(*
SPDX-FileCopyrightText: © 2026 Oleksandr Tiutyk <trofimich@gmail.com>
SPDX-License-Identifier: MIT
License: https://opensource.org/license/mit
*)

(*!
<summary>Describes typed generic storage and provides value access and conversion operations.</summary>
<description>
Stores a type category, address, byte size and ownership flag for externally stored data. Copying this
descriptor copies those fields, not the referenced payload. Typed access requires live storage matching the
descriptor; conversion methods do not validate its lifetime. Equals and GetHashCode share value semantics and
accept an optional borrowed IEqualityComparer. They preserve type categories, normalize floating NaN and
signed zero, and delegate nonempty OBJECT operands to the object's equality/hash pair. Neither method adds
descriptor state or takes ownership. Try methods contain exceptions and report failure without rolling back
bytes already written.
</description>
*)

{attribute 'no_explicit_call' := 'do not call this function block directly'}
FUNCTION_BLOCK GENERIC_VALUE
VAR_OUTPUT
	Address : POINTER TO BYTE;
	Size : ULINT;
	TypeClass : GENERIC_TYPE_CLASS;
	IsMemoryOwner : BOOL;
END_VAR

(*!
<summary>Returns a borrowed system descriptor for this generic value.</summary>
<description>
Does not copy the payload or transfer ownership. Size above SignedInt32.MAX_VALUE raises
ArgumentOutOfRangeException; type mapping exceptions propagate. The caller keeps the described storage alive
while using the result. Descendants cannot override this descriptor operation; customize value equality
through IEqualityComparer or the stored object equality contract.
</description>
*)
METHOD FINAL AsAnyType : __SYSTEM.AnyType
AsAnyType := SystemAnyTypes.CreateAnyTypeByGenericValue(genericValue := THIS^);
END_METHOD

(*!
<summary>Reads a Boolean or converts an integer to FALSE for zero and TRUE for any nonzero value.</summary>
<description>
Requires live storage matching the descriptor. Signed and unsigned integers are read at their full width,
including BYTE, WORD, DWORD and LWORD representations. Other categories throw
GenericConversionNotSupportedException. Stored data and ownership are unchanged. Descendants cannot override
this descriptor operation; customize value equality through IEqualityComparer or the stored object equality
contract.
</description>
*)
METHOD FINAL AsBool : BOOL
VAR
	universalPointer : UNIVERSAL_POINTER;
END_VAR
universalPointer.AsByte := Address;

CASE TypeClass OF
	GENERIC_TYPE_CLASS.BOOLEAN:
		AsBool := universalPointer.AsBool^;
		RETURN;

	GENERIC_TYPE_CLASS.INT_8, GENERIC_TYPE_CLASS.INT_16, GENERIC_TYPE_CLASS.INT_32, GENERIC_TYPE_CLASS.INT_64:
		AsBool := AsLInt() <> 0;
		RETURN;

	GENERIC_TYPE_CLASS.UINT_8, GENERIC_TYPE_CLASS.UINT_16, GENERIC_TYPE_CLASS.UINT_32, GENERIC_TYPE_CLASS.UINT_64:
		AsBool := AsULInt() <> 0;
		RETURN;
END_CASE

Exceptions.ThrowGenericConversionNotSupported(
		sourceNamespaceName := NamespaceName,
		sourceClassName := ClassName,
		sourcePOUName := __POUNAME(),
		sourcePosition := __POSITION(),
		sourceDataType := TypeClass,
		targetDataType := GENERIC_TYPE_CLASS.BOOLEAN
	);
END_METHOD

(*!
<summary>Reads or converts an integer representation when the value fits the result.</summary>
<description>
Requires live storage matching the descriptor. For supported integer types, FALSE accepts the actual value
only when it fits the result range; bounds are checked before narrowing or changing signedness. TRUE permits
the native conversion even outside that range. Unsupported types or rejected values raise
GenericConversionNotSupportedException. Existing BOOLEAN byte-view behavior is retained. Stored data and
ownership are unchanged; no dynamic allocation is needed for successful conversion. Descendants cannot
override this descriptor operation; customize value equality through IEqualityComparer or the stored object
equality contract.
</description>
*)
//!<param name="allowTypeCastWithDataLoss">
//! Allows native conversion when the actual value is outside the result range; overflow behavior follows
//! TwinCAT.
//! </param>
METHOD FINAL AsByte : BYTE
VAR_INPUT
	allowTypeCastWithDataLoss : BOOL := FALSE;
END_VAR
VAR
	universalPointer : UNIVERSAL_POINTER;
END_VAR
universalPointer.AsByte := Address;

CASE TypeClass OF
	GENERIC_TYPE_CLASS.BOOLEAN, GENERIC_TYPE_CLASS.UINT_8:
		 AsByte := universalPointer.AsByte^;
		 RETURN;

	GENERIC_TYPE_CLASS.UINT_16:
		IF allowTypeCastWithDataLoss OR_ELSE (TO_ULINT(universalPointer.AsWord^) <= TO_ULINT(UnsignedInt8.MAX_VALUE)) THEN
			AsByte := TO_BYTE(universalPointer.AsWord^);
			RETURN;
		END_IF

	GENERIC_TYPE_CLASS.UINT_32:
		IF allowTypeCastWithDataLoss OR_ELSE (TO_ULINT(universalPointer.AsDWord^) <= TO_ULINT(UnsignedInt8.MAX_VALUE)) THEN
			AsByte := TO_BYTE(universalPointer.AsDWord^);
			RETURN;
		END_IF

	GENERIC_TYPE_CLASS.UINT_64:
		IF allowTypeCastWithDataLoss OR_ELSE (TO_ULINT(universalPointer.AsLWord^) <= TO_ULINT(UnsignedInt8.MAX_VALUE)) THEN
			AsByte := TO_BYTE(universalPointer.AsLWord^);
			RETURN;
		END_IF

	GENERIC_TYPE_CLASS.INT_8:
		IF allowTypeCastWithDataLoss OR_ELSE (TO_LINT(universalPointer.AsSInt^) >= TO_LINT(UnsignedInt8.MIN_VALUE)) THEN
			AsByte := TO_BYTE(universalPointer.AsSInt^);
			RETURN;
		END_IF

	GENERIC_TYPE_CLASS.INT_16:
		IF allowTypeCastWithDataLoss
			OR_ELSE (TO_LINT(universalPointer.AsInt^) >= TO_LINT(UnsignedInt8.MIN_VALUE)
				AND_THEN TO_LINT(universalPointer.AsInt^) <= TO_LINT(UnsignedInt8.MAX_VALUE))
		THEN
			AsByte := TO_BYTE(universalPointer.AsInt^);
			RETURN;
		END_IF

	GENERIC_TYPE_CLASS.INT_32:
		IF allowTypeCastWithDataLoss
			OR_ELSE (TO_LINT(universalPointer.AsDInt^) >= TO_LINT(UnsignedInt8.MIN_VALUE)
				AND_THEN TO_LINT(universalPointer.AsDInt^) <= TO_LINT(UnsignedInt8.MAX_VALUE))
		THEN
			AsByte := TO_BYTE(universalPointer.AsDInt^);
			RETURN;
		END_IF

	GENERIC_TYPE_CLASS.INT_64:
		IF allowTypeCastWithDataLoss
			OR_ELSE (TO_LINT(universalPointer.AsLInt^) >= TO_LINT(UnsignedInt8.MIN_VALUE)
				AND_THEN TO_LINT(universalPointer.AsLInt^) <= TO_LINT(UnsignedInt8.MAX_VALUE))
		THEN
			AsByte := TO_BYTE(universalPointer.AsLInt^);
			RETURN;
		END_IF
END_CASE

Exceptions.ThrowGenericConversionNotSupported(
		sourceNamespaceName := NamespaceName,
		sourceClassName := ClassName,
		sourcePOUName := __POUNAME(),
		sourcePosition := __POSITION(),
		sourceDataType := TypeClass,
		targetDataType := GENERIC_TYPE_CLASS.UINT_8
	);
END_METHOD

(*!
<summary>Reads or converts a supported generic value to DATE.</summary>
<description>
Requires live storage matching the descriptor. INT_32, UINT_32, INT_64 and UINT_64 are counts of seconds since
the epoch; DATE_AND_TIME_32 is a calendar timestamp. Numeric inputs must fit DateAndTimes.MIN_VALUE/MAX_VALUE
even with TRUE. LDATE is checked as signed nanoseconds against the same limits widened to LDT before
narrowing. For these inputs, FALSE accepts only midnight; TRUE discards the time of day. The result of these
conversions has no hidden time remainder. Rejected or unsupported conversions raise
GenericConversionNotSupportedException. DATE_32 is read directly. A valid calendar LDATE within the DATE range
is accepted with either flag; a hidden time remainder requires TRUE and is explicitly removed. Stored data and
ownership are unchanged. Descendants cannot override this descriptor operation; customize value equality
through IEqualityComparer or the stored object equality contract.
</description>
*)
//!<param name="allowTypeCastWithDataLoss">
//! Allows discarding the time of day from numeric, DT and LDATE inputs; does not permit numeric or LDATE
//! range overflow.
//! </param>
METHOD FINAL AsDate : DATE
VAR_INPUT
	allowTypeCastWithDataLoss : BOOL := FALSE;
END_VAR
VAR
	universalPointer : UNIVERSAL_POINTER;

	secondsSinceMidnight : UDINT;
END_VAR
universalPointer.AsByte := Address;

CASE TypeClass OF
	GENERIC_TYPE_CLASS.DATE_32: 
		 AsDate := universalPointer.AsDate^;
		 RETURN;		 

	GENERIC_TYPE_CLASS.INT_32:
		IF universalPointer.AsDInt^ >= TO_LINT(DateAndTimes.MIN_VALUE) THEN
			secondsSinceMidnight := TO_UDINT(universalPointer.AsDInt^) MOD Times.SECONDS_PER_DAY;

			IF allowTypeCastWithDataLoss
				OR_ELSE secondsSinceMidnight = 0
			THEN
				AsDate := TO_DATE(TO_UDINT(universalPointer.AsDInt^) - secondsSinceMidnight);
				RETURN;
			END_IF
		END_IF

	GENERIC_TYPE_CLASS.UINT_32, GENERIC_TYPE_CLASS.DATE_AND_TIME_32:
		secondsSinceMidnight := TO_UDINT(universalPointer.AsUDInt^) MOD Times.SECONDS_PER_DAY;

		IF allowTypeCastWithDataLoss
			OR_ELSE secondsSinceMidnight = 0
		THEN
			AsDate := TO_DATE(TO_UDINT(universalPointer.AsUDInt^) - secondsSinceMidnight);
			RETURN;
		END_IF

	GENERIC_TYPE_CLASS.INT_64:
		IF universalPointer.AsLInt^ >= TO_LINT(DateAndTimes.MIN_VALUE) AND_THEN universalPointer.AsLInt^ <= TO_LINT(DateAndTimes.MAX_VALUE) THEN
			secondsSinceMidnight := TO_UDINT(universalPointer.AsLInt^) MOD Times.SECONDS_PER_DAY;

			IF allowTypeCastWithDataLoss
				OR_ELSE secondsSinceMidnight = 0
			THEN
				AsDate := TO_DATE(TO_UDINT(universalPointer.AsLInt^) - secondsSinceMidnight);
				RETURN;
			END_IF
		END_IF

	GENERIC_TYPE_CLASS.UINT_64:
		IF universalPointer.AsULInt^ <= TO_ULINT(DateAndTimes.MAX_VALUE) THEN
			secondsSinceMidnight := TO_UDINT(universalPointer.AsULInt^) MOD Times.SECONDS_PER_DAY;

			IF allowTypeCastWithDataLoss
				OR_ELSE secondsSinceMidnight = 0
			THEN
				AsDate := TO_DATE(TO_UDINT(universalPointer.AsULInt^) - secondsSinceMidnight);
				RETURN;
			END_IF
		END_IF

	GENERIC_TYPE_CLASS.DATE_64:
		IF universalPointer.AsLInt^ >= TO_LINT(TO_LDT(DateAndTimes.MIN_VALUE))
			AND_THEN universalPointer.AsLInt^ <= TO_LINT(TO_LDT(DateAndTimes.MAX_VALUE)) THEN
			IF allowTypeCastWithDataLoss OR_ELSE universalPointer.AsLInt^ MOD TO_LINT(LongTimes.ONE_DAY) = 0 THEN
				// Remove the time in nanoseconds before converting whole seconds to DATE.
				AsDate := TO_DATE((universalPointer.AsLInt^ - universalPointer.AsLInt^ MOD TO_LINT(LongTimes.ONE_DAY))
					/ TO_LINT(LongTimes.ONE_SECOND));
				RETURN;
			END_IF
		END_IF
END_CASE

Exceptions.ThrowGenericConversionNotSupported(
		sourceNamespaceName := NamespaceName,
		sourceClassName := ClassName,
		sourcePOUName := __POUNAME(),
		sourcePosition := __POSITION(),
		sourceDataType := TypeClass,
		targetDataType := GENERIC_TYPE_CLASS.DATE_32
	);
END_METHOD

(*!
<summary>Reads or converts a supported generic value to DATE_AND_TIME.</summary>
<description>
Requires live storage matching the descriptor. For DATE_AND_TIME_64, FALSE requires a timestamp within the DT
range and an exact whole number of seconds. Signed nanoseconds are checked before narrowing. TRUE uses native
TO_DT without these checks; out-of-range behavior depends on the runtime and may raise an exception. Rejected
or unsupported conversions raise GenericConversionNotSupportedException. Numeric inputs are seconds since the
epoch. With FALSE, signed inputs must be nonnegative and 64-bit inputs must fit the DT range; TRUE passes the
original signed or unsigned value to native TO_DT. DATE_32 and DATE_AND_TIME_32 retain their direct conversion
paths. Stored data and ownership are unchanged. Descendants cannot override this descriptor operation;
customize value equality through IEqualityComparer or the stored object equality contract.
</description>
*)
//!<param name="allowTypeCastWithDataLoss">
//! Allows loss of precision or range in LDT to DT conversion and native numeric conversions outside the DT
//! range.
//! </param>
METHOD FINAL AsDateAndTime : DATE_AND_TIME
VAR_INPUT
	allowTypeCastWithDataLoss : BOOL := FALSE;
END_VAR
VAR
	universalPointer : UNIVERSAL_POINTER;
END_VAR
universalPointer.AsByte := Address;

CASE TypeClass OF
	GENERIC_TYPE_CLASS.DATE_AND_TIME_32:
		 AsDateAndTime := universalPointer.AsDateAndTime^;
		 RETURN;

	GENERIC_TYPE_CLASS.UINT_32:
		 AsDateAndTime := TO_DT(universalPointer.AsUDInt^);
		 RETURN;
		
	GENERIC_TYPE_CLASS.DATE_32:
		 AsDateAndTime := TO_DT(universalPointer.AsDate^);
		 RETURN;
	GENERIC_TYPE_CLASS.DATE_AND_TIME_64:
		IF allowTypeCastWithDataLoss OR_ELSE (
			universalPointer.AsLInt^ >= TO_LINT(TO_LDT(DateAndTimes.MIN_VALUE))
			AND_THEN universalPointer.AsLInt^ <= TO_LINT(TO_LDT(DateAndTimes.MAX_VALUE))
			AND_THEN universalPointer.AsLInt^ MOD TO_LINT(LongTimes.ONE_SECOND) = 0) THEN
			AsDateAndTime := TO_DT(universalPointer.AsLDateAndTime^);
			RETURN;
		END_IF

	GENERIC_TYPE_CLASS.INT_32:
		IF allowTypeCastWithDataLoss OR_ELSE universalPointer.AsDInt^ >= TO_LINT(DateAndTimes.MIN_VALUE) THEN
			AsDateAndTime := TO_DT(universalPointer.AsDInt^);
			RETURN;
		END_IF

	GENERIC_TYPE_CLASS.INT_64:
		IF allowTypeCastWithDataLoss OR_ELSE (
			universalPointer.AsLInt^ >= TO_LINT(DateAndTimes.MIN_VALUE)
			AND_THEN universalPointer.AsLInt^ <= TO_LINT(DateAndTimes.MAX_VALUE)) THEN
			AsDateAndTime := TO_DT(universalPointer.AsLInt^);
			RETURN;
		END_IF

	GENERIC_TYPE_CLASS.UINT_64:
		IF allowTypeCastWithDataLoss OR_ELSE universalPointer.AsULInt^ <= TO_ULINT(DateAndTimes.MAX_VALUE) THEN
			AsDateAndTime := TO_DT(universalPointer.AsULInt^);
			RETURN;
		END_IF
END_CASE

Exceptions.ThrowGenericConversionNotSupported(
		sourceNamespaceName := NamespaceName,
		sourceClassName := ClassName,
		sourcePOUName := __POUNAME(),
		sourcePosition := __POSITION(),
		sourceDataType := TypeClass,
		targetDataType := GENERIC_TYPE_CLASS.DATE_AND_TIME_32
	);
END_METHOD

(*!
<summary>Reads or converts an integer representation when the value fits the result.</summary>
<description>
Requires live storage matching the descriptor. For supported integer types, FALSE accepts the actual value
only when it fits the result range; bounds are checked before narrowing or changing signedness. TRUE permits
the native conversion even outside that range. Unsupported types or rejected values raise
GenericConversionNotSupportedException. Existing BOOLEAN byte-view behavior is retained. Stored data and
ownership are unchanged; no dynamic allocation is needed for successful conversion. Descendants cannot
override this descriptor operation; customize value equality through IEqualityComparer or the stored object
equality contract.
</description>
*)
//!<param name="allowTypeCastWithDataLoss">
//! Allows native conversion when the actual value is outside the result range; overflow behavior follows
//! TwinCAT.
//! </param>
METHOD FINAL AsDInt : DINT
VAR_INPUT
	allowTypeCastWithDataLoss : BOOL := FALSE;
END_VAR
VAR
	universalPointer : UNIVERSAL_POINTER;
END_VAR
universalPointer.AsByte := Address;

CASE TypeClass OF
	GENERIC_TYPE_CLASS.BOOLEAN, GENERIC_TYPE_CLASS.UINT_8:
		 AsDInt := TO_DINT(universalPointer.AsByte^);
		 RETURN;
		
	GENERIC_TYPE_CLASS.UINT_16:
		 AsDInt := TO_DINT(universalPointer.AsWord^);
		 RETURN;

	GENERIC_TYPE_CLASS.INT_8: 
		 AsDInt := TO_DINT(universalPointer.AsSInt^);
		 RETURN;
		 
	GENERIC_TYPE_CLASS.INT_16: 
		 AsDInt := TO_DINT(universalPointer.AsInt^);
		 RETURN;
		 
	GENERIC_TYPE_CLASS.INT_32: 
		 AsDInt := universalPointer.AsDInt^;
		 RETURN;

	GENERIC_TYPE_CLASS.UINT_32:
		IF allowTypeCastWithDataLoss OR_ELSE (TO_ULINT(universalPointer.AsDWord^) <= TO_ULINT(SignedInt32.MAX_VALUE)) THEN
			AsDInt := TO_DINT(universalPointer.AsDWord^);
			RETURN;
		END_IF

	GENERIC_TYPE_CLASS.UINT_64:
		IF allowTypeCastWithDataLoss OR_ELSE (TO_ULINT(universalPointer.AsLWord^) <= TO_ULINT(SignedInt32.MAX_VALUE)) THEN
			AsDInt := TO_DINT(universalPointer.AsLWord^);
			RETURN;
		END_IF

	GENERIC_TYPE_CLASS.INT_64:
		IF allowTypeCastWithDataLoss
			OR_ELSE (TO_LINT(universalPointer.AsLInt^) >= TO_LINT(SignedInt32.MIN_VALUE)
				AND_THEN TO_LINT(universalPointer.AsLInt^) <= TO_LINT(SignedInt32.MAX_VALUE))
		THEN
			AsDInt := TO_DINT(universalPointer.AsLInt^);
			RETURN;
		END_IF
END_CASE

Exceptions.ThrowGenericConversionNotSupported(
		sourceNamespaceName := NamespaceName,
		sourceClassName := ClassName,
		sourcePOUName := __POUNAME(),
		sourcePosition := __POSITION(),
		sourceDataType := TypeClass,
		targetDataType := GENERIC_TYPE_CLASS.INT_32
	);
END_METHOD

(*!
<summary>Reads or converts an integer representation when the value fits the result.</summary>
<description>
Requires live storage matching the descriptor. For supported integer types, FALSE accepts the actual value
only when it fits the result range; bounds are checked before narrowing or changing signedness. TRUE permits
the native conversion even outside that range. Unsupported types or rejected values raise
GenericConversionNotSupportedException. Existing BOOLEAN byte-view behavior is retained. Stored data and
ownership are unchanged; no dynamic allocation is needed for successful conversion. Descendants cannot
override this descriptor operation; customize value equality through IEqualityComparer or the stored object
equality contract.
</description>
*)
//!<param name="allowTypeCastWithDataLoss">
//! Allows native conversion when the actual value is outside the result range; overflow behavior follows
//! TwinCAT.
//! </param>
METHOD FINAL AsDWord : DWORD
VAR_INPUT
	allowTypeCastWithDataLoss : BOOL := FALSE;
END_VAR
VAR
	universalPointer : UNIVERSAL_POINTER;
END_VAR
universalPointer.AsByte := Address;

CASE TypeClass OF
	GENERIC_TYPE_CLASS.BOOLEAN, GENERIC_TYPE_CLASS.UINT_8:
		 AsDWord := TO_DWORD(universalPointer.AsByte^);
		 RETURN;
		 
	GENERIC_TYPE_CLASS.UINT_16:
		 AsDWord := TO_DWORD(universalPointer.AsWord^);
		 RETURN;
 
	GENERIC_TYPE_CLASS.UINT_32: 
		 AsDWord := universalPointer.AsDWord^;
		 RETURN;

	GENERIC_TYPE_CLASS.UINT_64:
		IF allowTypeCastWithDataLoss OR_ELSE (TO_ULINT(universalPointer.AsLWord^) <= TO_ULINT(UnsignedInt32.MAX_VALUE)) THEN
			AsDWord := TO_DWORD(universalPointer.AsLWord^);
			RETURN;
		END_IF

	GENERIC_TYPE_CLASS.INT_8:
		IF allowTypeCastWithDataLoss OR_ELSE (TO_LINT(universalPointer.AsSInt^) >= TO_LINT(UnsignedInt32.MIN_VALUE)) THEN
			AsDWord := TO_DWORD(universalPointer.AsSInt^);
			RETURN;
		END_IF

	GENERIC_TYPE_CLASS.INT_16:
		IF allowTypeCastWithDataLoss OR_ELSE (TO_LINT(universalPointer.AsInt^) >= TO_LINT(UnsignedInt32.MIN_VALUE)) THEN
			AsDWord := TO_DWORD(universalPointer.AsInt^);
			RETURN;
		END_IF

	GENERIC_TYPE_CLASS.INT_32:
		IF allowTypeCastWithDataLoss OR_ELSE (TO_LINT(universalPointer.AsDInt^) >= TO_LINT(UnsignedInt32.MIN_VALUE)) THEN
			AsDWord := TO_DWORD(universalPointer.AsDInt^);
			RETURN;
		END_IF

	GENERIC_TYPE_CLASS.INT_64:
		IF allowTypeCastWithDataLoss
			OR_ELSE (TO_LINT(universalPointer.AsLInt^) >= TO_LINT(UnsignedInt32.MIN_VALUE)
				AND_THEN TO_LINT(universalPointer.AsLInt^) <= TO_LINT(UnsignedInt32.MAX_VALUE))
		THEN
			AsDWord := TO_DWORD(universalPointer.AsLInt^);
			RETURN;
		END_IF
END_CASE

Exceptions.ThrowGenericConversionNotSupported(
		sourceNamespaceName := NamespaceName,
		sourceClassName := ClassName,
		sourcePOUName := __POUNAME(),
		sourcePosition := __POSITION(),
		sourceDataType := TypeClass,
		targetDataType := GENERIC_TYPE_CLASS.UINT_32
	);
END_METHOD

(*!
<summary>Reads or converts an integer representation when the value fits the result.</summary>
<description>
Requires live storage matching the descriptor. For supported integer types, FALSE accepts the actual value
only when it fits the result range; bounds are checked before narrowing or changing signedness. TRUE permits
the native conversion even outside that range. Unsupported types or rejected values raise
GenericConversionNotSupportedException. Existing BOOLEAN byte-view behavior is retained. Stored data and
ownership are unchanged; no dynamic allocation is needed for successful conversion. Descendants cannot
override this descriptor operation; customize value equality through IEqualityComparer or the stored object
equality contract.
</description>
*)
//!<param name="allowTypeCastWithDataLoss">
//! Allows native conversion when the actual value is outside the result range; overflow behavior follows
//! TwinCAT.
//! </param>
METHOD FINAL AsInt : INT
VAR_INPUT
	allowTypeCastWithDataLoss : BOOL := FALSE;
END_VAR
VAR
	universalPointer : UNIVERSAL_POINTER;
END_VAR
universalPointer.AsByte := Address;

CASE TypeClass OF
	GENERIC_TYPE_CLASS.BOOLEAN, GENERIC_TYPE_CLASS.UINT_8:
		 AsInt := TO_INT(universalPointer.AsByte^);
		 RETURN;

	GENERIC_TYPE_CLASS.INT_8: 
		 AsInt := TO_INT(universalPointer.AsSInt^);
		 RETURN;
			 
	GENERIC_TYPE_CLASS.INT_16: 
		 AsInt := universalPointer.AsInt^;
		 RETURN;

	GENERIC_TYPE_CLASS.UINT_16:
		IF allowTypeCastWithDataLoss OR_ELSE (TO_ULINT(universalPointer.AsWord^) <= TO_ULINT(SignedInt16.MAX_VALUE)) THEN
			AsInt := TO_INT(universalPointer.AsWord^);
			RETURN;
		END_IF

	GENERIC_TYPE_CLASS.UINT_32:
		IF allowTypeCastWithDataLoss OR_ELSE (TO_ULINT(universalPointer.AsDWord^) <= TO_ULINT(SignedInt16.MAX_VALUE)) THEN
			AsInt := TO_INT(universalPointer.AsDWord^);
			RETURN;
		END_IF

	GENERIC_TYPE_CLASS.UINT_64:
		IF allowTypeCastWithDataLoss OR_ELSE (TO_ULINT(universalPointer.AsLWord^) <= TO_ULINT(SignedInt16.MAX_VALUE)) THEN
			AsInt := TO_INT(universalPointer.AsLWord^);
			RETURN;
		END_IF

	GENERIC_TYPE_CLASS.INT_32:
		IF allowTypeCastWithDataLoss
			OR_ELSE (TO_LINT(universalPointer.AsDInt^) >= TO_LINT(SignedInt16.MIN_VALUE)
				AND_THEN TO_LINT(universalPointer.AsDInt^) <= TO_LINT(SignedInt16.MAX_VALUE))
		THEN
			AsInt := TO_INT(universalPointer.AsDInt^);
			RETURN;
		END_IF

	GENERIC_TYPE_CLASS.INT_64:
		IF allowTypeCastWithDataLoss
			OR_ELSE (TO_LINT(universalPointer.AsLInt^) >= TO_LINT(SignedInt16.MIN_VALUE)
				AND_THEN TO_LINT(universalPointer.AsLInt^) <= TO_LINT(SignedInt16.MAX_VALUE))
		THEN
			AsInt := TO_INT(universalPointer.AsLInt^);
			RETURN;
		END_IF
END_CASE

Exceptions.ThrowGenericConversionNotSupported(
		sourceNamespaceName := NamespaceName,
		sourceClassName := ClassName,
		sourcePOUName := __POUNAME(),
		sourcePosition := __POSITION(),
		sourceDataType := TypeClass,
		targetDataType := GENERIC_TYPE_CLASS.INT_16
	);
END_METHOD

(*!
<summary>Returns a borrowed IObject view of object storage.</summary>
<description>
Requires OBJECT TypeClass; other tags raise GenericConversionNotSupportedException. A null address returns a
null interface; a nonnull address must identify a live compatible object. Does not clone or transfer
ownership. Descendants cannot override this descriptor operation; customize value equality through
IEqualityComparer or the stored object equality contract.
</description>
*)
METHOD FINAL AsIObject : IObject
VAR
	objectPointer : POINTER TO Object;

END_VAR
IF TypeClass = GENERIC_TYPE_CLASS.OBJECT THEN
	objectPointer := Address;
	
	IF objectPointer <> 0 THEN
		__QUERYINTERFACE(objectPointer^, AsIObject);						
	END_IF
ELSE	
	Exceptions.ThrowGenericConversionNotSupported(
		sourceNamespaceName := NamespaceName,
		sourceClassName := ClassName,
		sourcePOUName := __POUNAME(),
		sourcePosition := __POSITION(),
		sourceDataType := TypeClass,
		targetDataType := GENERIC_TYPE_CLASS.OBJECT
	);		
END_IF
END_METHOD

(*!
<summary>Reads or converts a supported generic value to LDATE.</summary>
<description>
Requires live storage matching the descriptor. DATE_AND_TIME_32 and DATE_AND_TIME_64 are treated as calendar
timestamps. INT_64 and UINT_64 are signed and unsigned counts of nanoseconds since the epoch. UINT_64 values
above LongDateAndTimes.MAX_VALUE are rejected even with TRUE. Numeric inputs follow calendar normalization:
FALSE accepts only midnight; TRUE discards the time of day. The results have no hidden time remainder. LDT
normalization uses signed nanoseconds and rounds down to midnight, including before the epoch. The first
partial LDT day (1677-09-21) is rejected even with TRUE because its midnight cannot be represented in LDATE;
the range check precedes subtraction. Rejected or unsupported conversions raise
GenericConversionNotSupportedException. DATE_64 is read directly and DATE_32 uses native widening; these paths
do not normalize hidden time components. Stored data and ownership are unchanged. Descendants cannot override
this descriptor operation; customize value equality through IEqualityComparer or the stored object equality
contract.
</description>
*)
//!<param name="allowTypeCastWithDataLoss">
//! Allows discarding the time of day from DT, LDT and numeric nanosecond counts; does not permit a midnight
//! outside the LDATE range.
//! </param>
METHOD FINAL AsLDate : LDATE
VAR_INPUT
	allowTypeCastWithDataLoss : BOOL := FALSE;
END_VAR
VAR
	universalPointer : UNIVERSAL_POINTER;

	secondsSinceMidnight : UDINT;
	nanosecondsSinceMidnight : LINT;
END_VAR
universalPointer.AsByte := Address;

CASE TypeClass OF
	GENERIC_TYPE_CLASS.DATE_64: 
		 AsLDate := universalPointer.AsLDate^;
		 RETURN;		 

	GENERIC_TYPE_CLASS.DATE_32: 
		 AsLDate := TO_LDATE(universalPointer.AsDate^);
		 RETURN;
	GENERIC_TYPE_CLASS.UINT_64:
		IF universalPointer.AsULInt^ <= TO_ULINT(LongDateAndTimes.MAX_VALUE) THEN
			nanosecondsSinceMidnight := TO_LINT(universalPointer.AsULInt^ MOD TO_ULINT(LongTimes.ONE_DAY));

			IF allowTypeCastWithDataLoss
				OR_ELSE nanosecondsSinceMidnight = 0
			THEN
				AsLDate := TO_LDATE(universalPointer.AsULInt^ - TO_ULINT(nanosecondsSinceMidnight));
				RETURN;
			END_IF
		END_IF

	GENERIC_TYPE_CLASS.DATE_AND_TIME_32:
		secondsSinceMidnight := TO_UDINT(universalPointer.AsDateAndTime^) MOD Times.SECONDS_PER_DAY;

		IF allowTypeCastWithDataLoss
			OR_ELSE secondsSinceMidnight = 0
		THEN
			AsLDate := TO_LDATE(TO_DT(TO_UDINT(universalPointer.AsDateAndTime^) - secondsSinceMidnight));
			RETURN;
		END_IF

	GENERIC_TYPE_CLASS.DATE_AND_TIME_64, GENERIC_TYPE_CLASS.INT_64:
		nanosecondsSinceMidnight := universalPointer.AsLInt^ MOD TO_LINT(LongTimes.ONE_DAY);

		// Normalize a negative remainder to the elapsed time since midnight.
		IF nanosecondsSinceMidnight < 0 THEN
			nanosecondsSinceMidnight := nanosecondsSinceMidnight + TO_LINT(LongTimes.ONE_DAY);
		END_IF

		IF (allowTypeCastWithDataLoss OR_ELSE nanosecondsSinceMidnight = 0)
			AND_THEN universalPointer.AsLInt^ >= SignedInt64.MIN_VALUE + nanosecondsSinceMidnight THEN
			AsLDate := TO_LDATE(universalPointer.AsLInt^ - nanosecondsSinceMidnight);
			RETURN;
		END_IF
END_CASE

Exceptions.ThrowGenericConversionNotSupported(
		sourceNamespaceName := NamespaceName,
		sourceClassName := ClassName,
		sourcePOUName := __POUNAME(),
		sourcePosition := __POSITION(),
		sourceDataType := TypeClass,
		targetDataType := GENERIC_TYPE_CLASS.DATE_64
	);
END_METHOD

(*!
<summary>Reads or converts a supported generic value to LDATE_AND_TIME.</summary>
<description>
Requires live storage matching the descriptor. Reads LDT directly and widens DT or DATE to LDT; valid LDATE is
also accepted with FALSE. Numeric INT_64 and UINT_64 inputs are nanoseconds since the epoch. INT_64 is read as
signed and fits the documented LDT range. UINT_64 with FALSE must not exceed LongDateAndTimes.MAX_VALUE; TRUE
permits native TO_LDT outside that range, with runtime-dependent results or exceptions. TIME and LTIME mean
duration added to the epoch. TIME milliseconds are scaled to nanoseconds in ULINT and always fit LDT. LTIME
already uses nanoseconds; FALSE checks LongDateAndTimes.MAX_VALUE before conversion, while TRUE allows native
out-of-range conversion. Rejected or unsupported conversions raise GenericConversionNotSupportedException.
Stored data and ownership are unchanged. Descendants cannot override this descriptor operation; customize
value equality through IEqualityComparer or the stored object equality contract.
</description>
*)
//!<param name="allowTypeCastWithDataLoss">Allows native out-of-range UINT_64 and LTIME conversion.</param>
METHOD FINAL AsLDateAndTime : LDATE_AND_TIME
VAR_INPUT
	allowTypeCastWithDataLoss : BOOL := FALSE;
END_VAR
VAR
	universalPointer : UNIVERSAL_POINTER;
END_VAR
universalPointer.AsByte := Address;

CASE TypeClass OF
	GENERIC_TYPE_CLASS.DATE_AND_TIME_64: 
		 AsLDateAndTime := universalPointer.AsLDateAndTime^;
		 RETURN;		 

	GENERIC_TYPE_CLASS.DATE_AND_TIME_32:
		 AsLDateAndTime := TO_LDT(universalPointer.AsDateAndTime^);
		 RETURN;
		 
	GENERIC_TYPE_CLASS.INT_64:
		AsLDateAndTime := TO_LDT(universalPointer.AsLInt^);
		RETURN;

	GENERIC_TYPE_CLASS.UINT_64:
		IF allowTypeCastWithDataLoss OR_ELSE universalPointer.AsULInt^ <= TO_ULINT(LongDateAndTimes.MAX_VALUE) THEN
			AsLDateAndTime := TO_LDT(universalPointer.AsULInt^);
			RETURN;
		END_IF

	GENERIC_TYPE_CLASS.DATE_32:
		 AsLDateAndTime := TO_LDT(universalPointer.AsDate^);
		 RETURN;

	GENERIC_TYPE_CLASS.TIME_32:
		 AsLDateAndTime := TO_LDT(TO_ULINT(universalPointer.AsTime^) * TO_ULINT(LongTimes.ONE_MILLISECOND));
		 RETURN;
	GENERIC_TYPE_CLASS.DATE_64:
		AsLDateAndTime := TO_LDT(universalPointer.AsLDate^);
		RETURN;

	GENERIC_TYPE_CLASS.TIME_64:
		IF allowTypeCastWithDataLoss OR_ELSE TO_ULINT(universalPointer.AsLTime^) <= TO_ULINT(LongDateAndTimes.MAX_VALUE) THEN
			AsLDateAndTime := TO_LDT(TO_ULINT(universalPointer.AsLTime^));
			RETURN;
		END_IF
END_CASE

Exceptions.ThrowGenericConversionNotSupported(
		sourceNamespaceName := NamespaceName,
		sourceClassName := ClassName,
		sourcePOUName := __POUNAME(),
		sourcePosition := __POSITION(),
		sourceDataType := TypeClass,
		targetDataType := GENERIC_TYPE_CLASS.DATE_AND_TIME_64
	);
END_METHOD

(*!
<summary>Reads or converts an integer representation when the value fits the result.</summary>
<description>
Requires live storage matching the descriptor. For supported integer types, FALSE accepts the actual value
only when it fits the result range; bounds are checked before narrowing or changing signedness. TRUE permits
the native conversion even outside that range. Unsupported types or rejected values raise
GenericConversionNotSupportedException. Existing BOOLEAN byte-view behavior is retained. Stored data and
ownership are unchanged; no dynamic allocation is needed for successful conversion. Descendants cannot
override this descriptor operation; customize value equality through IEqualityComparer or the stored object
equality contract.
</description>
*)
//!<param name="allowTypeCastWithDataLoss">
//! Allows native conversion when the actual value is outside the result range; overflow behavior follows
//! TwinCAT.
//! </param>
METHOD FINAL AsLInt : LINT
VAR_INPUT
	allowTypeCastWithDataLoss : BOOL := FALSE;
END_VAR
VAR
	universalPointer : UNIVERSAL_POINTER;
END_VAR
universalPointer.AsByte := Address;

CASE TypeClass OF
	GENERIC_TYPE_CLASS.BOOLEAN, GENERIC_TYPE_CLASS.UINT_8:
		 AsLInt := TO_LINT(universalPointer.AsByte^);
		 RETURN;
		
	GENERIC_TYPE_CLASS.UINT_16:
		 AsLInt := TO_LINT(universalPointer.AsWord^);
		 RETURN;

	GENERIC_TYPE_CLASS.UINT_32: 
		 AsLInt := TO_LINT(universalPointer.AsDWord^);
		 RETURN;

	GENERIC_TYPE_CLASS.INT_8: 
		 AsLInt := TO_LINT(universalPointer.AsSInt^);
		 RETURN;
		 
	GENERIC_TYPE_CLASS.INT_16: 
		 AsLInt := TO_LINT(universalPointer.AsInt^);
		 RETURN;
		 
	GENERIC_TYPE_CLASS.INT_32: 
		 AsLInt := TO_LINT(universalPointer.AsDInt^);
		 RETURN;
			 			 
	GENERIC_TYPE_CLASS.INT_64:
		 AsLInt := universalPointer.AsLInt^;
		 RETURN;

	GENERIC_TYPE_CLASS.UINT_64:
		IF allowTypeCastWithDataLoss OR_ELSE (TO_ULINT(universalPointer.AsLWord^) <= TO_ULINT(SignedInt64.MAX_VALUE)) THEN
			AsLInt := TO_LINT(universalPointer.AsLWord^);
			RETURN;
		END_IF
END_CASE

Exceptions.ThrowGenericConversionNotSupported(
		sourceNamespaceName := NamespaceName,
		sourceClassName := ClassName,
		sourcePOUName := __POUNAME(),
		sourcePosition := __POSITION(),
		sourceDataType := TypeClass,
		targetDataType := GENERIC_TYPE_CLASS.INT_64
	);
END_METHOD

(*!
<summary>Reads REAL_32 or REAL_64 storage as LREAL.</summary>
<description>
REAL_32 is widened and REAL_64 read directly. Other tags raise GenericConversionNotSupportedException. The
address must reference live, aligned storage of the tagged representation. Descendants cannot override this
descriptor operation; customize value equality through IEqualityComparer or the stored object equality
contract.
</description>
*)
METHOD FINAL AsLReal : LREAL
VAR
	universalPointer : UNIVERSAL_POINTER;
END_VAR
universalPointer.AsByte := Address;

CASE TypeClass OF
	GENERIC_TYPE_CLASS.BOOLEAN, GENERIC_TYPE_CLASS.UINT_8:
		AsLReal := TO_LREAL(universalPointer.AsByte^);
		RETURN;

	GENERIC_TYPE_CLASS.UINT_16:
		AsLReal := TO_LREAL(universalPointer.AsWord^);
		RETURN;

	GENERIC_TYPE_CLASS.UINT_32:
		AsLReal := TO_LREAL(universalPointer.AsDWord^);
		RETURN;

	GENERIC_TYPE_CLASS.UINT_64:
		AsLReal := TO_LREAL(universalPointer.AsLWord^);
		RETURN;

	GENERIC_TYPE_CLASS.INT_8:
		AsLReal := TO_LREAL(universalPointer.AsSInt^);
		RETURN;

	GENERIC_TYPE_CLASS.INT_16:
		AsLReal := TO_LREAL(universalPointer.AsInt^);
		RETURN;

	GENERIC_TYPE_CLASS.INT_32:
		AsLReal := TO_LREAL(universalPointer.AsDInt^);
		RETURN;

	GENERIC_TYPE_CLASS.INT_64:
		AsLReal := TO_LREAL(universalPointer.AsLInt^);
		RETURN;

	GENERIC_TYPE_CLASS.REAL_32:
		AsLReal := TO_LREAL(universalPointer.AsReal^);
		RETURN;
	 
	GENERIC_TYPE_CLASS.REAL_64:	
		AsLReal := universalPointer.AsLReal^;
		RETURN;
END_CASE

Exceptions.ThrowGenericConversionNotSupported(
		sourceNamespaceName := NamespaceName,
		sourceClassName := ClassName,
		sourcePOUName := __POUNAME(),
		sourcePosition := __POSITION(),
		sourceDataType := TypeClass,
		targetDataType := GENERIC_TYPE_CLASS.REAL_64
	);
END_METHOD

(*!
<summary>Reads or converts a supported generic value to a nanosecond duration.</summary>
<description>
Requires live storage matching the descriptor. DT and LDT inputs mean elapsed time since the epoch. DT seconds
are scaled to nanoseconds in ULINT and always fit LTIME. LDT is read as signed nanoseconds; FALSE rejects
timestamps before the epoch, while TRUE passes the signed value to native TO_LTIME. INT_64 follows the same
nonnegative rule. Valid TOD/LTOD inputs mean duration since midnight. TIME_32 is widened; TIME_64 and UINT_64
retain their values. TRUE does not guarantee safe out-of-range behavior. Unsupported or rejected conversions
raise GenericConversionNotSupportedException. Stored data and ownership are unchanged. Descendants cannot
override this descriptor operation; customize value equality through IEqualityComparer or the stored object
equality contract.
</description>
*)
//!<param name="allowTypeCastWithDataLoss">
//! Allows native conversion of negative INT_64 values and LDT timestamps before the epoch.
//! </param>
METHOD FINAL AsLTime : LTIME
VAR_INPUT
	allowTypeCastWithDataLoss : BOOL := FALSE;
END_VAR
VAR
	universalPointer : UNIVERSAL_POINTER;
END_VAR
universalPointer.AsByte := Address;

CASE TypeClass OF
	GENERIC_TYPE_CLASS.TIME_64:
		 AsLTime := universalPointer.AsLTime^;
		 RETURN;

	GENERIC_TYPE_CLASS.TIME_32: 
		 AsLTime := TO_LTIME(universalPointer.AsTime^);
		 RETURN;
		
	GENERIC_TYPE_CLASS.UINT_64:
		 AsLTime := TO_LTIME(universalPointer.AsULInt^);
		 RETURN;

	GENERIC_TYPE_CLASS.DATE_AND_TIME_32:
		 AsLTime := TO_LTIME(TO_ULINT(universalPointer.AsDateAndTime^) * TO_ULINT(LongTimes.ONE_SECOND));
		 RETURN;
		 
	GENERIC_TYPE_CLASS.TIME_OF_DAY_32: 
		 AsLTime := TO_LTIME(universalPointer.AsTimeOfDay^);
		 RETURN;

	GENERIC_TYPE_CLASS.TIME_OF_DAY_64:
		AsLTime := TO_LTIME(universalPointer.AsLTimeOfDay^);
		RETURN;

	GENERIC_TYPE_CLASS.INT_64:
		IF allowTypeCastWithDataLoss OR_ELSE universalPointer.AsLInt^ >= TO_LINT(LongTimes.MIN_VALUE) THEN
			AsLTime := TO_LTIME(universalPointer.AsLInt^);
			RETURN;
		END_IF

	GENERIC_TYPE_CLASS.DATE_AND_TIME_64:
		IF allowTypeCastWithDataLoss OR_ELSE universalPointer.AsLInt^ >= TO_LINT(LongDateAndTimes.EPOCH) THEN
			AsLTime := TO_LTIME(universalPointer.AsLInt^);
			RETURN;
		END_IF
END_CASE

Exceptions.ThrowGenericConversionNotSupported(
		sourceNamespaceName := NamespaceName,
		sourceClassName := ClassName,
		sourcePOUName := __POUNAME(),
		sourcePosition := __POSITION(),
		sourceDataType := TypeClass,
		targetDataType := GENERIC_TYPE_CLASS.TIME_64
	);
END_METHOD

(*!
<summary>Reads or converts a supported generic value to LTIME_OF_DAY.</summary>
<description>
Reads a time of day in nanoseconds. With FALSE, supported integer and duration inputs must be nonnegative and
less than 24 hours; integer units are nanoseconds. TIME_OF_DAY_64 is read directly and TIME_OF_DAY_32 is
widened. TRUE permits out-of-range native conversions. For DT/LDT, FALSE accepts only timestamps on
1970-01-01; TRUE discards the calendar date and extracts the time of day. Negative LDT remainders are
normalized to the interval from midnight inclusive to one day exclusive. Nanosecond precision is preserved.
Requires live storage matching the descriptor. Checks precede the potentially lossy conversion. Rejected or
unsupported conversions raise GenericConversionNotSupportedException. TRUE does not guarantee safe overflow
behavior. Stored data and ownership are unchanged. Descendants cannot override this descriptor operation;
customize value equality through IEqualityComparer or the stored object equality contract.
</description>
*)
//!<param name="allowTypeCastWithDataLoss">
//! Allows native conversion when the value cannot be represented exactly; FALSE checks numeric and duration
//! inputs and rejects DT/LDT dates other than 1970-01-01.
//! </param>
METHOD FINAL AsLTimeOfDay : LTIME_OF_DAY
VAR_INPUT
	allowTypeCastWithDataLoss : BOOL := FALSE;
END_VAR
VAR
	universalPointer : UNIVERSAL_POINTER;

	nanosecondsSinceMidnight : LINT;
END_VAR
universalPointer.AsByte := Address;

CASE TypeClass OF
	GENERIC_TYPE_CLASS.TIME_OF_DAY_64:
		AsLTimeOfDay := universalPointer.AsLTimeOfDay^;
		RETURN;

	GENERIC_TYPE_CLASS.TIME_OF_DAY_32:
		AsLTimeOfDay := TO_LTOD(universalPointer.AsTimeOfDay^);
		RETURN;

	GENERIC_TYPE_CLASS.UINT_64:
		IF allowTypeCastWithDataLoss OR_ELSE (universalPointer.AsULInt^ < TO_ULINT(LongTimes.ONE_DAY)) THEN
			AsLTimeOfDay := TO_LTOD(universalPointer.AsULInt^);
			RETURN;
		END_IF

	GENERIC_TYPE_CLASS.INT_64:
		IF allowTypeCastWithDataLoss
			OR_ELSE (universalPointer.AsLInt^ >= TO_LINT(LongTimes.MIN_VALUE) AND_THEN universalPointer.AsLInt^ < TO_LINT(LongTimes.ONE_DAY))
		THEN
			AsLTimeOfDay := TO_LTOD(universalPointer.AsLInt^);
			RETURN;
		END_IF

	GENERIC_TYPE_CLASS.TIME_32:
		IF allowTypeCastWithDataLoss
			OR_ELSE (universalPointer.AsTime^ < Times.ONE_DAY)
		THEN
			AsLTimeOfDay := TO_LTOD(universalPointer.AsTime^);
			RETURN;
		END_IF

	GENERIC_TYPE_CLASS.DATE_AND_TIME_32:
		IF allowTypeCastWithDataLoss OR_ELSE TO_UDINT(universalPointer.AsDateAndTime^) < Times.SECONDS_PER_DAY THEN
			AsLTimeOfDay := TO_LTOD(TO_ULINT(TO_UDINT(universalPointer.AsDateAndTime^) MOD Times.SECONDS_PER_DAY)
				* TO_ULINT(LongTimes.ONE_SECOND));
			RETURN;
		END_IF

	GENERIC_TYPE_CLASS.TIME_64:
		IF allowTypeCastWithDataLoss
			OR_ELSE (universalPointer.AsLTime^ < LongTimes.ONE_DAY)
		THEN
			AsLTimeOfDay := TO_LTOD(universalPointer.AsLTime^);
			RETURN;
		END_IF

	GENERIC_TYPE_CLASS.DATE_AND_TIME_64:
		IF allowTypeCastWithDataLoss OR_ELSE (
			universalPointer.AsLInt^ >= TO_LINT(LongDateAndTimes.EPOCH)
			AND_THEN universalPointer.AsLInt^ < TO_LINT(LongTimes.ONE_DAY)) THEN
			nanosecondsSinceMidnight := universalPointer.AsLInt^ MOD TO_LINT(LongTimes.ONE_DAY);

			IF nanosecondsSinceMidnight < 0 THEN
				nanosecondsSinceMidnight := nanosecondsSinceMidnight + TO_LINT(LongTimes.ONE_DAY);
			END_IF

			AsLTimeOfDay := TO_LTOD(nanosecondsSinceMidnight);
			RETURN;
		END_IF

END_CASE

Exceptions.ThrowGenericConversionNotSupported(
		sourceNamespaceName := NamespaceName,
		sourceClassName := ClassName,
		sourcePOUName := __POUNAME(),
		sourcePosition := __POSITION(),
		sourceDataType := TypeClass,
		targetDataType := GENERIC_TYPE_CLASS.TIME_OF_DAY_64
	);
END_METHOD

(*!
<summary>Reads or converts an integer representation when the value fits the result.</summary>
<description>
Requires live storage matching the descriptor. For supported integer types, FALSE accepts the actual value
only when it fits the result range; bounds are checked before narrowing or changing signedness. TRUE permits
the native conversion even outside that range. Unsupported types or rejected values raise
GenericConversionNotSupportedException. Existing BOOLEAN byte-view behavior is retained. Stored data and
ownership are unchanged; no dynamic allocation is needed for successful conversion. Descendants cannot
override this descriptor operation; customize value equality through IEqualityComparer or the stored object
equality contract.
</description>
*)
//!<param name="allowTypeCastWithDataLoss">
//! Allows native conversion when the actual value is outside the result range; overflow behavior follows
//! TwinCAT.
//! </param>
METHOD FINAL AsLWord : LWORD
VAR_INPUT
	allowTypeCastWithDataLoss : BOOL := FALSE;
END_VAR
VAR
	universalPointer : UNIVERSAL_POINTER;
END_VAR
universalPointer.AsByte := Address;

CASE TypeClass OF
	GENERIC_TYPE_CLASS.BOOLEAN, GENERIC_TYPE_CLASS.UINT_8:
		 AsLWord := TO_LWORD(universalPointer.AsByte^);
		 RETURN;
		 
	GENERIC_TYPE_CLASS.UINT_16:
		 AsLWord := TO_LWORD(universalPointer.AsWord^);
		 RETURN;
 
	GENERIC_TYPE_CLASS.UINT_32: 
		 AsLWord := TO_LWORD(universalPointer.AsDWord^);
		 RETURN;
		 
	GENERIC_TYPE_CLASS.UINT_64:	
		 AsLWord := universalPointer.AsLWord^;
		 RETURN;

	GENERIC_TYPE_CLASS.INT_8:
		IF allowTypeCastWithDataLoss OR_ELSE (TO_LINT(universalPointer.AsSInt^) >= TO_LINT(UnsignedInt64.MIN_VALUE)) THEN
			AsLWord := TO_LWORD(universalPointer.AsSInt^);
			RETURN;
		END_IF

	GENERIC_TYPE_CLASS.INT_16:
		IF allowTypeCastWithDataLoss OR_ELSE (TO_LINT(universalPointer.AsInt^) >= TO_LINT(UnsignedInt64.MIN_VALUE)) THEN
			AsLWord := TO_LWORD(universalPointer.AsInt^);
			RETURN;
		END_IF

	GENERIC_TYPE_CLASS.INT_32:
		IF allowTypeCastWithDataLoss OR_ELSE (TO_LINT(universalPointer.AsDInt^) >= TO_LINT(UnsignedInt64.MIN_VALUE)) THEN
			AsLWord := TO_LWORD(universalPointer.AsDInt^);
			RETURN;
		END_IF

	GENERIC_TYPE_CLASS.INT_64:
		IF allowTypeCastWithDataLoss OR_ELSE (TO_LINT(universalPointer.AsLInt^) >= TO_LINT(UnsignedInt64.MIN_VALUE)) THEN
			AsLWord := TO_LWORD(universalPointer.AsLInt^);
			RETURN;
		END_IF
END_CASE

Exceptions.ThrowGenericConversionNotSupported(
		sourceNamespaceName := NamespaceName,
		sourceClassName := ClassName,
		sourcePOUName := __POUNAME(),
		sourcePosition := __POSITION(),
		sourceDataType := TypeClass,
		targetDataType := GENERIC_TYPE_CLASS.UINT_64
	);
END_METHOD

(*!
<summary>Returns a borrowed reference to object storage.</summary>
<description>
Requires OBJECT TypeClass; other tags raise GenericConversionNotSupportedException. A null address leaves the
result unbound. A nonnull address must identify a live Object; the reference does not extend its lifetime.
Descendants cannot override this descriptor operation; customize value equality through IEqualityComparer or
the stored object equality contract.
</description>
*)
METHOD FINAL AsObject : REFERENCE TO Object
VAR
	objectPointer : POINTER TO Object;

END_VAR
IF TypeClass = GENERIC_TYPE_CLASS.OBJECT THEN
	objectPointer := Address;
	
	IF objectPointer <> 0 THEN
		AsObject REF= objectPointer^;		
	END_IF
ELSE	
	Exceptions.ThrowGenericConversionNotSupported(
		sourceNamespaceName := NamespaceName,
		sourceClassName := ClassName,
		sourcePOUName := __POUNAME(),
		sourcePosition := __POSITION(),
		sourceDataType := TypeClass,
		targetDataType := GENERIC_TYPE_CLASS.OBJECT
	);		
END_IF
END_METHOD

(*!
<summary>Reads a REAL value or converts an LREAL value according to its representability.</summary>
<description>
Requires live storage matching TypeClass. REAL_32 is read directly. For REAL_64 with FALSE, rejects NaN and
infinities by their exponent bits, checks the finite REAL range before narrowing, and accepts the result only
if widening it back to LREAL reproduces the original value. With TRUE, uses native TO_REAL without these
checks, including for special values. Native floating-point behavior follows the target runtime configuration.
Unsupported or inexact conversions with FALSE raise GenericConversionNotSupportedException. Stored data and
ownership are unchanged. Descendants cannot override this descriptor operation; customize value equality
through IEqualityComparer or the stored object equality contract.
</description>
*)
//!<param name="allowTypeCastWithDataLoss">
//! Allows inexact, out-of-range and special-value LREAL to REAL conversions; FALSE requires a finite exactly
//! representable value.
//! </param>
METHOD FINAL AsReal : REAL
VAR_INPUT
	allowTypeCastWithDataLoss : BOOL := FALSE;
END_VAR
VAR
	universalPointer : UNIVERSAL_POINTER;
END_VAR
universalPointer.AsByte := Address;

CASE TypeClass OF
	GENERIC_TYPE_CLASS.REAL_32:
		AsReal := universalPointer.AsReal^;
		RETURN;

	GENERIC_TYPE_CLASS.REAL_64:
		IF allowTypeCastWithDataLoss THEN
			AsReal := TO_REAL(universalPointer.AsLReal^);
			RETURN;
		END_IF

		// All exponent bits are set for both infinity and NaN.
		IF (universalPointer.AsULInt^ AND LongReals.POSITIVE_INFINITY.Raw) <> LongReals.POSITIVE_INFINITY.Raw
			AND_THEN universalPointer.AsLReal^ >= TO_LREAL(Reals.MIN_VALUE)
			AND_THEN universalPointer.AsLReal^ <= TO_LREAL(Reals.MAX_VALUE) THEN
			AsReal := TO_REAL(universalPointer.AsLReal^);

			IF TO_LREAL(AsReal) = universalPointer.AsLReal^ THEN
				RETURN;
			END_IF
		END_IF
END_CASE

Exceptions.ThrowGenericConversionNotSupported(
		sourceNamespaceName := NamespaceName,
		sourceClassName := ClassName,
		sourcePOUName := __POUNAME(),
		sourcePosition := __POSITION(),
		sourceDataType := TypeClass,
		targetDataType := GENERIC_TYPE_CLASS.REAL_32
	);
END_METHOD

(*!
<summary>Installs descriptor fields without copying or releasing a payload.</summary>
<description>
A null address raises ArgumentNotSpecifiedException before modification. The caller supplies a consistent
type, size and ownership flag and must arrange release of any previous owned storage before overwriting it.
Descendants cannot override this descriptor operation; customize value equality through IEqualityComparer or
the stored object equality contract.
</description>
*)
METHOD INTERNAL FINAL Assign
VAR_INPUT
	genericTypeClass : GENERIC_TYPE_CLASS;
	address : POINTER TO BYTE;
	size : ULINT;
	isMemoryOwner : BOOL;
END_VAR
IF address = 0 THEN
	Exceptions.ThrowArgumentNotSpecified(
		sourceNamespaceName := NamespaceName,
		sourceClassName := ClassName,
		sourcePOUName := __POUNAME(),
		sourcePosition := __POSITION(),
		argumentName := 'address'
	);
END_IF

THIS^.TypeClass := genericTypeClass;
THIS^.Address := address;
THIS^.Size := size;
THIS^.IsMemoryOwner := isMemoryOwner;
END_METHOD

(*!
<summary>Reads or converts an integer representation when the value fits the result.</summary>
<description>
Requires live storage matching the descriptor. For supported integer types, FALSE accepts the actual value
only when it fits the result range; bounds are checked before narrowing or changing signedness. TRUE permits
the native conversion even outside that range. Unsupported types or rejected values raise
GenericConversionNotSupportedException. Existing BOOLEAN byte-view behavior is retained. Stored data and
ownership are unchanged; no dynamic allocation is needed for successful conversion. Descendants cannot
override this descriptor operation; customize value equality through IEqualityComparer or the stored object
equality contract.
</description>
*)
//!<param name="allowTypeCastWithDataLoss">
//! Allows native conversion when the actual value is outside the result range; overflow behavior follows
//! TwinCAT.
//! </param>
METHOD FINAL AsSInt : SINT
VAR_INPUT
	allowTypeCastWithDataLoss : BOOL := FALSE;
END_VAR
VAR
	universalPointer : UNIVERSAL_POINTER;
END_VAR
universalPointer.AsByte := Address;

CASE TypeClass OF
	GENERIC_TYPE_CLASS.INT_8: 
		 AsSInt := universalPointer.AsSInt^;
		 RETURN;

	GENERIC_TYPE_CLASS.UINT_16:
		IF allowTypeCastWithDataLoss OR_ELSE (TO_ULINT(universalPointer.AsWord^) <= TO_ULINT(SignedInt8.MAX_VALUE)) THEN
			AsSInt := TO_SINT(universalPointer.AsWord^);
			RETURN;
		END_IF

	GENERIC_TYPE_CLASS.UINT_32:
		IF allowTypeCastWithDataLoss OR_ELSE (TO_ULINT(universalPointer.AsDWord^) <= TO_ULINT(SignedInt8.MAX_VALUE)) THEN
			AsSInt := TO_SINT(universalPointer.AsDWord^);
			RETURN;
		END_IF

	GENERIC_TYPE_CLASS.UINT_64:
		IF allowTypeCastWithDataLoss OR_ELSE (TO_ULINT(universalPointer.AsLWord^) <= TO_ULINT(SignedInt8.MAX_VALUE)) THEN
			AsSInt := TO_SINT(universalPointer.AsLWord^);
			RETURN;
		END_IF

	GENERIC_TYPE_CLASS.INT_16:
		IF allowTypeCastWithDataLoss
			OR_ELSE (TO_LINT(universalPointer.AsInt^) >= TO_LINT(SignedInt8.MIN_VALUE)
				AND_THEN TO_LINT(universalPointer.AsInt^) <= TO_LINT(SignedInt8.MAX_VALUE))
		THEN
			AsSInt := TO_SINT(universalPointer.AsInt^);
			RETURN;
		END_IF

	GENERIC_TYPE_CLASS.INT_32:
		IF allowTypeCastWithDataLoss
			OR_ELSE (TO_LINT(universalPointer.AsDInt^) >= TO_LINT(SignedInt8.MIN_VALUE)
				AND_THEN TO_LINT(universalPointer.AsDInt^) <= TO_LINT(SignedInt8.MAX_VALUE))
		THEN
			AsSInt := TO_SINT(universalPointer.AsDInt^);
			RETURN;
		END_IF

	GENERIC_TYPE_CLASS.INT_64:
		IF allowTypeCastWithDataLoss
			OR_ELSE (TO_LINT(universalPointer.AsLInt^) >= TO_LINT(SignedInt8.MIN_VALUE)
				AND_THEN TO_LINT(universalPointer.AsLInt^) <= TO_LINT(SignedInt8.MAX_VALUE))
		THEN
			AsSInt := TO_SINT(universalPointer.AsLInt^);
			RETURN;
		END_IF
END_CASE

Exceptions.ThrowGenericConversionNotSupported(
		sourceNamespaceName := NamespaceName,
		sourceClassName := ClassName,
		sourcePOUName := __POUNAME(),
		sourcePosition := __POSITION(),
		sourceDataType := TypeClass,
		targetDataType := GENERIC_TYPE_CLASS.INT_8
	);
END_METHOD

(*!
<summary>Formats a supported generic value as text with capacity for 255 characters.</summary>
<description>
Requires live storage matching the descriptor. Same-encoding string values are copied directly into the
result, retaining at most 255 code units and a terminator without an intermediate 80-character string. WSTRING
uses single-byte Latin-1 conversion, not UTF-8. With FALSE, each source code unit in the retained prefix (at
most 255, stopping at the terminator) must fit UnsignedByte.MAX_VALUE; otherwise
GenericConversionNotSupportedException is raised before conversion. The truncated tail is not validated. TRUE
permits omission of unrepresentable characters. WSTRING_TO_STRING2 writes directly into the result and skips
characters it cannot convert. Output beyond the 255-byte text capacity is not retained; the function
completion flag is intentionally ignored because this API permits truncation. Numeric formatting retains its
native conversion behavior. Unsupported conversions raise GenericConversionNotSupportedException; the source
and ownership are unchanged. Descendants cannot override this descriptor operation; customize value equality
through IEqualityComparer or the stored object equality contract.
</description>
*)
//!<param name="allowTypeCastWithDataLoss">
//! Allows omission of WSTRING characters that cannot be represented in Latin-1. Truncation to 255 bytes is
//! allowed with either flag.
//! </param>
METHOD FINAL AsString255 : STRING(255)
VAR_INPUT
	allowTypeCastWithDataLoss : BOOL := FALSE;
END_VAR
VAR
	universalPointer : UNIVERSAL_POINTER;

	characterIndex : UDINT;
END_VAR
universalPointer.AsByte := Address;

CASE TypeClass OF
	GENERIC_TYPE_CLASS.BOOLEAN:
		 AsString255 := TO_STRING(universalPointer.AsBool^);
		 RETURN;
    GENERIC_TYPE_CLASS.INT_8:
		 AsString255 := TO_STRING(universalPointer.AsSInt^);
		 RETURN;
    GENERIC_TYPE_CLASS.INT_16:
		 AsString255 := TO_STRING(universalPointer.AsInt^);
		 RETURN;
    GENERIC_TYPE_CLASS.INT_32:
		 AsString255 := TO_STRING(universalPointer.AsDInt^);
		 RETURN;
    GENERIC_TYPE_CLASS.INT_64:
		 AsString255 := TO_STRING(universalPointer.AsLInt^);
		 RETURN;
    GENERIC_TYPE_CLASS.UINT_8:
		 AsString255 := TO_STRING(universalPointer.AsUSInt^);
		 RETURN;
    GENERIC_TYPE_CLASS.UINT_16:
		 AsString255 := TO_STRING(universalPointer.AsUInt^);
		 RETURN;
    GENERIC_TYPE_CLASS.UINT_32:
		 AsString255 := TO_STRING(universalPointer.AsUDInt^);
		 RETURN;
    GENERIC_TYPE_CLASS.UINT_64:
		 AsString255 := TO_STRING(universalPointer.AsULInt^);
		 RETURN;
    GENERIC_TYPE_CLASS.REAL_32:
		 AsString255 := TO_STRING(universalPointer.AsReal^);
		 RETURN;
    GENERIC_TYPE_CLASS.REAL_64:
		 AsString255 := TO_STRING(universalPointer.AsLReal^);
		 RETURN;
    GENERIC_TYPE_CLASS.STRING_8:
		Tc2_Utilities.STRNCPY(
			pDst := ADR(AsString255),
			pSrc := universalPointer.AsString,
			nDstSize := SIZEOF(AsString255)
		);
		 RETURN;
    GENERIC_TYPE_CLASS.TIME_32:
		 AsString255 := TO_STRING(universalPointer.AsTime^);
		 RETURN;
    GENERIC_TYPE_CLASS.TIME_64:
		 AsString255 := TO_STRING(universalPointer.AsLTime^);
		 RETURN;
    GENERIC_TYPE_CLASS.DATE_32:
		 AsString255 := TO_STRING(universalPointer.AsDate^);
		 RETURN;
    GENERIC_TYPE_CLASS.DATE_64:
		 AsString255 := TO_STRING(universalPointer.AsLDate ^);
		 RETURN;
    GENERIC_TYPE_CLASS.DATE_AND_TIME_32:
		 AsString255 := TO_STRING(universalPointer.AsDateAndTime^);
		 RETURN;
    GENERIC_TYPE_CLASS.DATE_AND_TIME_64:
		 AsString255 := TO_STRING(universalPointer.AsLDateAndTime^);
		 RETURN;
    GENERIC_TYPE_CLASS.TIME_OF_DAY_32:
		 AsString255 := TO_STRING(universalPointer.AsTimeOfDay^);
		 RETURN;
    GENERIC_TYPE_CLASS.TIME_OF_DAY_64:
		 AsString255 := TO_STRING(universalPointer.AsLTimeOfDay^);
		 RETURN;

	GENERIC_TYPE_CLASS.STRING_16:
		IF NOT allowTypeCastWithDataLoss THEN
			FOR characterIndex := 0 TO SIZEOF(AsString255) - 2 DO
				IF universalPointer.AsWord[characterIndex] = 0 THEN
					EXIT;
				END_IF

				IF universalPointer.AsWord[characterIndex] > TO_WORD(UnsignedInt8.MAX_VALUE) THEN
					Exceptions.ThrowGenericConversionNotSupported(
						sourceNamespaceName := NamespaceName,
						sourceClassName := ClassName,
						sourcePOUName := __POUNAME(),
						sourcePosition := __POSITION(),
						sourceDataType := TypeClass,
		targetDataType := GENERIC_TYPE_CLASS.STRING_8
					);
				END_IF
			END_FOR
		END_IF

		Tc2_Utilities.WSTRING_TO_STRING2(
	pDstString := ADR(AsString255),
	pSrcWString := universalPointer.AsWString,
	nDstSize := SIZEOF(AsString255)
);
		RETURN;
END_CASE

Exceptions.ThrowGenericConversionNotSupported(
		sourceNamespaceName := NamespaceName,
		sourceClassName := ClassName,
		sourcePOUName := __POUNAME(),
		sourcePosition := __POSITION(),
		sourceDataType := TypeClass,
		targetDataType := GENERIC_TYPE_CLASS.STRING_8
	);
END_METHOD

(*!
<summary>Borrows the STRING storage described by this value.</summary>
<description>
Requires STRING_8 or raises GenericConversionNotSupportedException. Does not copy, bound-check or validate
the payload. The reference remains valid only while the source storage remains alive; the descriptor size
still limits any access. Descendants cannot override this descriptor operation; customize value equality
through IEqualityComparer or the stored object equality contract.
</description>
*)
METHOD FINAL AsStringReference : REFERENCE TO STRING
VAR
	universalPointer : UNIVERSAL_POINTER;
END_VAR
universalPointer.AsByte := Address;

CASE TypeClass OF
    GENERIC_TYPE_CLASS.STRING_8:
		 AsStringReference REF= universalPointer.AsString^;
		 RETURN;
END_CASE

Exceptions.ThrowGenericConversionNotSupported(
		sourceNamespaceName := NamespaceName,
		sourceClassName := ClassName,
		sourcePOUName := __POUNAME(),
		sourcePosition := __POSITION(),
		sourceDataType := TypeClass,
		targetDataType := GENERIC_TYPE_CLASS.STRING_8
	);
END_METHOD

(*!
<summary>Reads or converts a supported value to a millisecond duration.</summary>
<description>
DT input means elapsed time since the epoch: seconds are scaled to milliseconds in ULINT before conversion.
FALSE requires that duration to fit Times.MAX_VALUE; TRUE permits native out-of-range narrowing. Reads a
millisecond duration. With FALSE, signed integer inputs must be nonnegative and 64-bit integer inputs must fit
UINT_32; integer units are milliseconds. LTIME additionally must fit TIME and contain an integral number of
milliseconds. TRUE permits the native conversion even when these conditions fail. Requires live storage
matching the descriptor. Checks precede the potentially lossy conversion. Rejected or unsupported conversions
raise GenericConversionNotSupportedException. TRUE does not guarantee safe overflow behavior. Stored data and
ownership are unchanged. Descendants cannot override this descriptor operation; customize value equality
through IEqualityComparer or the stored object equality contract.
</description>
*)
//!<param name="allowTypeCastWithDataLoss">
//! Allows native conversion when the value cannot be represented exactly; FALSE checks supported numeric and
//! duration inputs.
//! </param>
METHOD FINAL AsTime : TIME
VAR_INPUT
	allowTypeCastWithDataLoss : BOOL := FALSE;
END_VAR
VAR
	universalPointer : UNIVERSAL_POINTER;
END_VAR
universalPointer.AsByte := Address;

CASE TypeClass OF
	GENERIC_TYPE_CLASS.DATE_AND_TIME_32:
		IF allowTypeCastWithDataLoss
			OR_ELSE TO_ULINT(universalPointer.AsDateAndTime^) <= TO_ULINT(Times.MAX_VALUE) / TO_ULINT(Times.ONE_SECOND)
		THEN
			AsTime := TO_TIME(TO_ULINT(universalPointer.AsDateAndTime^) * TO_ULINT(Times.ONE_SECOND));
			RETURN;
		END_IF

	GENERIC_TYPE_CLASS.UINT_32:
		AsTime := TO_TIME(universalPointer.AsUDInt^);
		RETURN;

	GENERIC_TYPE_CLASS.INT_32:
		IF allowTypeCastWithDataLoss OR_ELSE (universalPointer.AsDInt^ >= TO_LINT(Times.MIN_VALUE)) THEN
			AsTime := TO_TIME(universalPointer.AsDInt^);
			RETURN;
		END_IF

	GENERIC_TYPE_CLASS.TIME_32:
		AsTime := universalPointer.AsTime^;
		RETURN;

	GENERIC_TYPE_CLASS.TIME_OF_DAY_32:
		AsTime := TO_TIME(universalPointer.AsTimeOfDay^);
		RETURN;

	GENERIC_TYPE_CLASS.TIME_64:
		IF allowTypeCastWithDataLoss
			OR_ELSE (universalPointer.AsLTime^ <= TO_LTIME(Times.MAX_VALUE)
				AND_THEN TO_ULINT(universalPointer.AsLTime^) MOD TO_ULINT(LongTimes.ONE_MILLISECOND) = 0)
		THEN
			AsTime := TO_TIME(universalPointer.AsLTime^);
			RETURN;
		END_IF

	GENERIC_TYPE_CLASS.INT_64:
		IF allowTypeCastWithDataLoss
			OR_ELSE (universalPointer.AsLInt^ >= TO_LINT(Times.MIN_VALUE) AND_THEN universalPointer.AsLInt^ <= TO_LINT(Times.MAX_VALUE))
		THEN
			AsTime := TO_TIME(universalPointer.AsLInt^);
			RETURN;
		END_IF

	GENERIC_TYPE_CLASS.UINT_64:
		IF allowTypeCastWithDataLoss OR_ELSE (universalPointer.AsULInt^ <= TO_ULINT(Times.MAX_VALUE)) THEN
			AsTime := TO_TIME(universalPointer.AsULInt^);
			RETURN;
		END_IF

END_CASE

Exceptions.ThrowGenericConversionNotSupported(
		sourceNamespaceName := NamespaceName,
		sourceClassName := ClassName,
		sourcePOUName := __POUNAME(),
		sourcePosition := __POSITION(),
		sourceDataType := TypeClass,
		targetDataType := GENERIC_TYPE_CLASS.TIME_32
	);
END_METHOD

(*!
<summary>Reads or converts a supported generic value to TIME_OF_DAY.</summary>
<description>
Reads a time of day in milliseconds. With FALSE, supported integer and duration inputs must be nonnegative and
less than 24 hours; integer units are milliseconds. LTIME additionally must contain an integral number of
milliseconds. TRUE permits the native conversion even when these conditions fail. TIME_OF_DAY_32 is read
directly. Requires live storage matching the descriptor. Checks precede the potentially lossy conversion.
Rejected or unsupported conversions raise GenericConversionNotSupportedException. TRUE does not guarantee safe
overflow behavior. Stored data and ownership are unchanged. Descendants cannot override this descriptor
operation; customize value equality through IEqualityComparer or the stored object equality contract.
</description>
*)
//!<param name="allowTypeCastWithDataLoss">
//! Allows native conversion when the value cannot be represented exactly; FALSE checks supported numeric and
//! duration inputs.
//! </param>
METHOD FINAL AsTimeOfDay : TIME_OF_DAY
VAR_INPUT
	allowTypeCastWithDataLoss : BOOL := FALSE;
END_VAR
VAR
	universalPointer : UNIVERSAL_POINTER;
END_VAR
universalPointer.AsByte := Address;

CASE TypeClass OF
	GENERIC_TYPE_CLASS.TIME_OF_DAY_32:
		AsTimeOfDay := universalPointer.AsTimeOfDay^;
		RETURN;

	GENERIC_TYPE_CLASS.INT_32:
		IF allowTypeCastWithDataLoss
			OR_ELSE (universalPointer.AsDInt^ >= TO_LINT(Times.MIN_VALUE) AND_THEN universalPointer.AsDInt^ < TO_DINT(Times.ONE_DAY))
		THEN
			AsTimeOfDay := TO_TOD(universalPointer.AsDInt^);
			RETURN;
		END_IF

	GENERIC_TYPE_CLASS.UINT_32:
		IF allowTypeCastWithDataLoss OR_ELSE (universalPointer.AsUDInt^ < TO_UDINT(Times.ONE_DAY)) THEN
			AsTimeOfDay := TO_TOD(universalPointer.AsUDInt^);
			RETURN;
		END_IF

	GENERIC_TYPE_CLASS.TIME_32:
		IF allowTypeCastWithDataLoss
			OR_ELSE (universalPointer.AsTime^ < Times.ONE_DAY)
		THEN
			AsTimeOfDay := TO_TOD(universalPointer.AsTime^);
			RETURN;
		END_IF

	GENERIC_TYPE_CLASS.INT_64:
		IF allowTypeCastWithDataLoss
			OR_ELSE (universalPointer.AsLInt^ >= TO_LINT(Times.MIN_VALUE) AND_THEN universalPointer.AsLInt^ < TO_LINT(Times.ONE_DAY))
		THEN
			AsTimeOfDay := TO_TOD(universalPointer.AsLInt^);
			RETURN;
		END_IF

	GENERIC_TYPE_CLASS.UINT_64:
		IF allowTypeCastWithDataLoss OR_ELSE (universalPointer.AsULInt^ < TO_ULINT(Times.ONE_DAY)) THEN
			AsTimeOfDay := TO_TOD(universalPointer.AsULInt^);
			RETURN;
		END_IF

	GENERIC_TYPE_CLASS.TIME_64:
		IF allowTypeCastWithDataLoss
			OR_ELSE (universalPointer.AsLTime^ < LongTimes.ONE_DAY
				AND_THEN TO_ULINT(universalPointer.AsLTime^) MOD TO_ULINT(LongTimes.ONE_MILLISECOND) = 0)
		THEN
			AsTimeOfDay := TO_TOD(universalPointer.AsLTime^);
			RETURN;
		END_IF

END_CASE

Exceptions.ThrowGenericConversionNotSupported(
		sourceNamespaceName := NamespaceName,
		sourceClassName := ClassName,
		sourcePOUName := __POUNAME(),
		sourcePosition := __POSITION(),
		sourceDataType := TypeClass,
		targetDataType := GENERIC_TYPE_CLASS.TIME_OF_DAY_32
	);
END_METHOD

(*!
<summary>Reads or converts an integer representation when the value fits the result.</summary>
<description>
Requires live storage matching the descriptor. For supported integer types, FALSE accepts the actual value
only when it fits the result range; bounds are checked before narrowing or changing signedness. TRUE permits
the native conversion even outside that range. Unsupported types or rejected values raise
GenericConversionNotSupportedException. Existing BOOLEAN byte-view behavior is retained. Stored data and
ownership are unchanged; no dynamic allocation is needed for successful conversion. Descendants cannot
override this descriptor operation; customize value equality through IEqualityComparer or the stored object
equality contract.
</description>
*)
//!<param name="allowTypeCastWithDataLoss">
//! Allows native conversion when the actual value is outside the result range; overflow behavior follows
//! TwinCAT.
//! </param>
METHOD FINAL AsUDInt : UDINT
VAR_INPUT
	allowTypeCastWithDataLoss : BOOL := FALSE;
END_VAR
VAR
	universalPointer : UNIVERSAL_POINTER;
END_VAR
universalPointer.AsByte := Address;

CASE TypeClass OF
	GENERIC_TYPE_CLASS.BOOLEAN, GENERIC_TYPE_CLASS.UINT_8:
		 AsUDInt := TO_UDINT(universalPointer.AsByte^);
		 RETURN;
		 
	GENERIC_TYPE_CLASS.UINT_16:
		 AsUDInt := TO_UDINT(universalPointer.AsWord^);
		 RETURN;
 
	GENERIC_TYPE_CLASS.UINT_32: 
		 AsUDInt := universalPointer.AsDWord^;
		 RETURN;

	GENERIC_TYPE_CLASS.UINT_64:
		IF allowTypeCastWithDataLoss OR_ELSE (TO_ULINT(universalPointer.AsLWord^) <= TO_ULINT(UnsignedInt32.MAX_VALUE)) THEN
			AsUDInt := TO_UDINT(universalPointer.AsLWord^);
			RETURN;
		END_IF

	GENERIC_TYPE_CLASS.INT_8:
		IF allowTypeCastWithDataLoss OR_ELSE (TO_LINT(universalPointer.AsSInt^) >= TO_LINT(UnsignedInt32.MIN_VALUE)) THEN
			AsUDInt := TO_UDINT(universalPointer.AsSInt^);
			RETURN;
		END_IF

	GENERIC_TYPE_CLASS.INT_16:
		IF allowTypeCastWithDataLoss OR_ELSE (TO_LINT(universalPointer.AsInt^) >= TO_LINT(UnsignedInt32.MIN_VALUE)) THEN
			AsUDInt := TO_UDINT(universalPointer.AsInt^);
			RETURN;
		END_IF

	GENERIC_TYPE_CLASS.INT_32:
		IF allowTypeCastWithDataLoss OR_ELSE (TO_LINT(universalPointer.AsDInt^) >= TO_LINT(UnsignedInt32.MIN_VALUE)) THEN
			AsUDInt := TO_UDINT(universalPointer.AsDInt^);
			RETURN;
		END_IF

	GENERIC_TYPE_CLASS.INT_64:
		IF allowTypeCastWithDataLoss
			OR_ELSE (TO_LINT(universalPointer.AsLInt^) >= TO_LINT(UnsignedInt32.MIN_VALUE)
				AND_THEN TO_LINT(universalPointer.AsLInt^) <= TO_LINT(UnsignedInt32.MAX_VALUE))
		THEN
			AsUDInt := TO_UDINT(universalPointer.AsLInt^);
			RETURN;
		END_IF
END_CASE

Exceptions.ThrowGenericConversionNotSupported(
		sourceNamespaceName := NamespaceName,
		sourceClassName := ClassName,
		sourcePOUName := __POUNAME(),
		sourcePosition := __POSITION(),
		sourceDataType := TypeClass,
		targetDataType := GENERIC_TYPE_CLASS.UINT_32
	);
END_METHOD

(*!
<summary>Reads or converts an integer representation when the value fits the result.</summary>
<description>
Requires live storage matching the descriptor. For supported integer types, FALSE accepts the actual value
only when it fits the result range; bounds are checked before narrowing or changing signedness. TRUE permits
the native conversion even outside that range. Unsupported types or rejected values raise
GenericConversionNotSupportedException. Existing BOOLEAN byte-view behavior is retained. Stored data and
ownership are unchanged; no dynamic allocation is needed for successful conversion. Descendants cannot
override this descriptor operation; customize value equality through IEqualityComparer or the stored object
equality contract.
</description>
*)
//!<param name="allowTypeCastWithDataLoss">
//! Allows native conversion when the actual value is outside the result range; overflow behavior follows
//! TwinCAT.
//! </param>
METHOD FINAL AsUInt : UINT
VAR_INPUT
	allowTypeCastWithDataLoss : BOOL := FALSE;
END_VAR
VAR
	universalPointer : UNIVERSAL_POINTER;
END_VAR
universalPointer.AsByte := Address;

CASE TypeClass OF
	GENERIC_TYPE_CLASS.BOOLEAN, GENERIC_TYPE_CLASS.UINT_8:
		 AsUInt := TO_UINT(universalPointer.AsByte^);
		 RETURN;
		 
	GENERIC_TYPE_CLASS.UINT_16:
		 AsUInt := universalPointer.AsWord^;
		 RETURN;

	GENERIC_TYPE_CLASS.UINT_32:
		IF allowTypeCastWithDataLoss OR_ELSE (TO_ULINT(universalPointer.AsDWord^) <= TO_ULINT(UnsignedInt16.MAX_VALUE)) THEN
			AsUInt := TO_UINT(universalPointer.AsDWord^);
			RETURN;
		END_IF

	GENERIC_TYPE_CLASS.UINT_64:
		IF allowTypeCastWithDataLoss OR_ELSE (TO_ULINT(universalPointer.AsLWord^) <= TO_ULINT(UnsignedInt16.MAX_VALUE)) THEN
			AsUInt := TO_UINT(universalPointer.AsLWord^);
			RETURN;
		END_IF

	GENERIC_TYPE_CLASS.INT_8:
		IF allowTypeCastWithDataLoss OR_ELSE (TO_LINT(universalPointer.AsSInt^) >= TO_LINT(UnsignedInt16.MIN_VALUE)) THEN
			AsUInt := TO_UINT(universalPointer.AsSInt^);
			RETURN;
		END_IF

	GENERIC_TYPE_CLASS.INT_16:
		IF allowTypeCastWithDataLoss OR_ELSE (TO_LINT(universalPointer.AsInt^) >= TO_LINT(UnsignedInt16.MIN_VALUE)) THEN
			AsUInt := TO_UINT(universalPointer.AsInt^);
			RETURN;
		END_IF

	GENERIC_TYPE_CLASS.INT_32:
		IF allowTypeCastWithDataLoss
			OR_ELSE (TO_LINT(universalPointer.AsDInt^) >= TO_LINT(UnsignedInt16.MIN_VALUE)
				AND_THEN TO_LINT(universalPointer.AsDInt^) <= TO_LINT(UnsignedInt16.MAX_VALUE))
		THEN
			AsUInt := TO_UINT(universalPointer.AsDInt^);
			RETURN;
		END_IF

	GENERIC_TYPE_CLASS.INT_64:
		IF allowTypeCastWithDataLoss
			OR_ELSE (TO_LINT(universalPointer.AsLInt^) >= TO_LINT(UnsignedInt16.MIN_VALUE)
				AND_THEN TO_LINT(universalPointer.AsLInt^) <= TO_LINT(UnsignedInt16.MAX_VALUE))
		THEN
			AsUInt := TO_UINT(universalPointer.AsLInt^);
			RETURN;
		END_IF
END_CASE

Exceptions.ThrowGenericConversionNotSupported(
		sourceNamespaceName := NamespaceName,
		sourceClassName := ClassName,
		sourcePOUName := __POUNAME(),
		sourcePosition := __POSITION(),
		sourceDataType := TypeClass,
		targetDataType := GENERIC_TYPE_CLASS.UINT_16
	);
END_METHOD

(*!
<summary>Reads or converts an integer representation when the value fits the result.</summary>
<description>
Requires live storage matching the descriptor. For supported integer types, FALSE accepts the actual value
only when it fits the result range; bounds are checked before narrowing or changing signedness. TRUE permits
the native conversion even outside that range. Unsupported types or rejected values raise
GenericConversionNotSupportedException. Existing BOOLEAN byte-view behavior is retained. Stored data and
ownership are unchanged; no dynamic allocation is needed for successful conversion. Descendants cannot
override this descriptor operation; customize value equality through IEqualityComparer or the stored object
equality contract.
</description>
*)
//!<param name="allowTypeCastWithDataLoss">
//! Allows native conversion when the actual value is outside the result range; overflow behavior follows
//! TwinCAT.
//! </param>
METHOD FINAL AsULInt : ULINT
VAR_INPUT
	allowTypeCastWithDataLoss : BOOL := FALSE;
END_VAR
VAR
	universalPointer : UNIVERSAL_POINTER;
END_VAR
universalPointer.AsByte := Address;

CASE TypeClass OF
	GENERIC_TYPE_CLASS.BOOLEAN, GENERIC_TYPE_CLASS.UINT_8:
		 AsULInt := TO_ULINT(universalPointer.AsByte^);
		 RETURN;
		 
	GENERIC_TYPE_CLASS.UINT_16:
		 AsULInt := TO_ULINT(universalPointer.AsWord^);
		 RETURN;
 
	GENERIC_TYPE_CLASS.UINT_32: 
		 AsULInt := TO_ULINT(universalPointer.AsDWord^);
		 RETURN;
		 
	GENERIC_TYPE_CLASS.UINT_64:	
		 AsULInt := universalPointer.AsLWord^;
		 RETURN;

	GENERIC_TYPE_CLASS.INT_8:
		IF allowTypeCastWithDataLoss OR_ELSE (TO_LINT(universalPointer.AsSInt^) >= TO_LINT(UnsignedInt64.MIN_VALUE)) THEN
			AsULInt := TO_ULINT(universalPointer.AsSInt^);
			RETURN;
		END_IF

	GENERIC_TYPE_CLASS.INT_16:
		IF allowTypeCastWithDataLoss OR_ELSE (TO_LINT(universalPointer.AsInt^) >= TO_LINT(UnsignedInt64.MIN_VALUE)) THEN
			AsULInt := TO_ULINT(universalPointer.AsInt^);
			RETURN;
		END_IF

	GENERIC_TYPE_CLASS.INT_32:
		IF allowTypeCastWithDataLoss OR_ELSE (TO_LINT(universalPointer.AsDInt^) >= TO_LINT(UnsignedInt64.MIN_VALUE)) THEN
			AsULInt := TO_ULINT(universalPointer.AsDInt^);
			RETURN;
		END_IF

	GENERIC_TYPE_CLASS.INT_64:
		IF allowTypeCastWithDataLoss OR_ELSE (TO_LINT(universalPointer.AsLInt^) >= TO_LINT(UnsignedInt64.MIN_VALUE)) THEN
			AsULInt := TO_ULINT(universalPointer.AsLInt^);
			RETURN;
		END_IF
END_CASE

Exceptions.ThrowGenericConversionNotSupported(
		sourceNamespaceName := NamespaceName,
		sourceClassName := ClassName,
		sourcePOUName := __POUNAME(),
		sourcePosition := __POSITION(),
		sourceDataType := TypeClass,
		targetDataType := GENERIC_TYPE_CLASS.UINT_64
	);
END_METHOD

(*!
<summary>Reads or converts an integer representation when the value fits the result.</summary>
<description>
Requires live storage matching the descriptor. For supported integer types, FALSE accepts the actual value
only when it fits the result range; bounds are checked before narrowing or changing signedness. TRUE permits
the native conversion even outside that range. Unsupported types or rejected values raise
GenericConversionNotSupportedException. Existing BOOLEAN byte-view behavior is retained. Stored data and
ownership are unchanged; no dynamic allocation is needed for successful conversion. Descendants cannot
override this descriptor operation; customize value equality through IEqualityComparer or the stored object
equality contract.
</description>
*)
//!<param name="allowTypeCastWithDataLoss">
//! Allows native conversion when the actual value is outside the result range; overflow behavior follows
//! TwinCAT.
//! </param>
METHOD FINAL AsUSInt : USINT
VAR_INPUT
	allowTypeCastWithDataLoss : BOOL := FALSE;
END_VAR
VAR
	universalPointer : UNIVERSAL_POINTER;
END_VAR
universalPointer.AsByte := Address;

CASE TypeClass OF
	GENERIC_TYPE_CLASS.BOOLEAN, GENERIC_TYPE_CLASS.UINT_8:
		 AsUSInt := universalPointer.AsUSInt^;
		 RETURN;

	GENERIC_TYPE_CLASS.UINT_16:
		IF allowTypeCastWithDataLoss OR_ELSE (TO_ULINT(universalPointer.AsWord^) <= TO_ULINT(UnsignedInt8.MAX_VALUE)) THEN
			AsUSInt := TO_USINT(universalPointer.AsWord^);
			RETURN;
		END_IF

	GENERIC_TYPE_CLASS.UINT_32:
		IF allowTypeCastWithDataLoss OR_ELSE (TO_ULINT(universalPointer.AsDWord^) <= TO_ULINT(UnsignedInt8.MAX_VALUE)) THEN
			AsUSInt := TO_USINT(universalPointer.AsDWord^);
			RETURN;
		END_IF

	GENERIC_TYPE_CLASS.UINT_64:
		IF allowTypeCastWithDataLoss OR_ELSE (TO_ULINT(universalPointer.AsLWord^) <= TO_ULINT(UnsignedInt8.MAX_VALUE)) THEN
			AsUSInt := TO_USINT(universalPointer.AsLWord^);
			RETURN;
		END_IF

	GENERIC_TYPE_CLASS.INT_8:
		IF allowTypeCastWithDataLoss OR_ELSE (TO_LINT(universalPointer.AsSInt^) >= TO_LINT(UnsignedInt8.MIN_VALUE)) THEN
			AsUSInt := TO_USINT(universalPointer.AsSInt^);
			RETURN;
		END_IF

	GENERIC_TYPE_CLASS.INT_16:
		IF allowTypeCastWithDataLoss
			OR_ELSE (TO_LINT(universalPointer.AsInt^) >= TO_LINT(UnsignedInt8.MIN_VALUE)
				AND_THEN TO_LINT(universalPointer.AsInt^) <= TO_LINT(UnsignedInt8.MAX_VALUE))
		THEN
			AsUSInt := TO_USINT(universalPointer.AsInt^);
			RETURN;
		END_IF

	GENERIC_TYPE_CLASS.INT_32:
		IF allowTypeCastWithDataLoss
			OR_ELSE (TO_LINT(universalPointer.AsDInt^) >= TO_LINT(UnsignedInt8.MIN_VALUE)
				AND_THEN TO_LINT(universalPointer.AsDInt^) <= TO_LINT(UnsignedInt8.MAX_VALUE))
		THEN
			AsUSInt := TO_USINT(universalPointer.AsDInt^);
			RETURN;
		END_IF

	GENERIC_TYPE_CLASS.INT_64:
		IF allowTypeCastWithDataLoss
			OR_ELSE (TO_LINT(universalPointer.AsLInt^) >= TO_LINT(UnsignedInt8.MIN_VALUE)
				AND_THEN TO_LINT(universalPointer.AsLInt^) <= TO_LINT(UnsignedInt8.MAX_VALUE))
		THEN
			AsUSInt := TO_USINT(universalPointer.AsLInt^);
			RETURN;
		END_IF
END_CASE

Exceptions.ThrowGenericConversionNotSupported(
		sourceNamespaceName := NamespaceName,
		sourceClassName := ClassName,
		sourcePOUName := __POUNAME(),
		sourcePosition := __POSITION(),
		sourceDataType := TypeClass,
		targetDataType := GENERIC_TYPE_CLASS.UINT_8
	);
END_METHOD

(*!
<summary>Reads or converts an integer representation when the value fits the result.</summary>
<description>
Requires live storage matching the descriptor. For supported integer types, FALSE accepts the actual value
only when it fits the result range; bounds are checked before narrowing or changing signedness. TRUE permits
the native conversion even outside that range. Unsupported types or rejected values raise
GenericConversionNotSupportedException. Existing BOOLEAN byte-view behavior is retained. Stored data and
ownership are unchanged; no dynamic allocation is needed for successful conversion. Descendants cannot
override this descriptor operation; customize value equality through IEqualityComparer or the stored object
equality contract.
</description>
*)
//!<param name="allowTypeCastWithDataLoss">
//! Allows native conversion when the actual value is outside the result range; overflow behavior follows
//! TwinCAT.
//! </param>
METHOD FINAL AsWord : WORD
VAR_INPUT
	allowTypeCastWithDataLoss : BOOL := FALSE;
END_VAR
VAR
	universalPointer : UNIVERSAL_POINTER;
END_VAR
universalPointer.AsByte := Address;

CASE TypeClass OF
	GENERIC_TYPE_CLASS.BOOLEAN, GENERIC_TYPE_CLASS.UINT_8:
		 AsWord := TO_WORD(universalPointer.AsByte^);
		 RETURN;
		 
	GENERIC_TYPE_CLASS.UINT_16:
		 AsWord := universalPointer.AsWord^;
		 RETURN;

	GENERIC_TYPE_CLASS.UINT_32:
		IF allowTypeCastWithDataLoss OR_ELSE (TO_ULINT(universalPointer.AsDWord^) <= TO_ULINT(UnsignedInt16.MAX_VALUE)) THEN
			AsWord := TO_WORD(universalPointer.AsDWord^);
			RETURN;
		END_IF

	GENERIC_TYPE_CLASS.UINT_64:
		IF allowTypeCastWithDataLoss OR_ELSE (TO_ULINT(universalPointer.AsLWord^) <= TO_ULINT(UnsignedInt16.MAX_VALUE)) THEN
			AsWord := TO_WORD(universalPointer.AsLWord^);
			RETURN;
		END_IF

	GENERIC_TYPE_CLASS.INT_8:
		IF allowTypeCastWithDataLoss OR_ELSE (TO_LINT(universalPointer.AsSInt^) >= TO_LINT(UnsignedInt16.MIN_VALUE)) THEN
			AsWord := TO_WORD(universalPointer.AsSInt^);
			RETURN;
		END_IF

	GENERIC_TYPE_CLASS.INT_16:
		IF allowTypeCastWithDataLoss OR_ELSE (TO_LINT(universalPointer.AsInt^) >= TO_LINT(UnsignedInt16.MIN_VALUE)) THEN
			AsWord := TO_WORD(universalPointer.AsInt^);
			RETURN;
		END_IF

	GENERIC_TYPE_CLASS.INT_32:
		IF allowTypeCastWithDataLoss
			OR_ELSE (TO_LINT(universalPointer.AsDInt^) >= TO_LINT(UnsignedInt16.MIN_VALUE)
				AND_THEN TO_LINT(universalPointer.AsDInt^) <= TO_LINT(UnsignedInt16.MAX_VALUE))
		THEN
			AsWord := TO_WORD(universalPointer.AsDInt^);
			RETURN;
		END_IF

	GENERIC_TYPE_CLASS.INT_64:
		IF allowTypeCastWithDataLoss
			OR_ELSE (TO_LINT(universalPointer.AsLInt^) >= TO_LINT(UnsignedInt16.MIN_VALUE)
				AND_THEN TO_LINT(universalPointer.AsLInt^) <= TO_LINT(UnsignedInt16.MAX_VALUE))
		THEN
			AsWord := TO_WORD(universalPointer.AsLInt^);
			RETURN;
		END_IF
END_CASE

Exceptions.ThrowGenericConversionNotSupported(
		sourceNamespaceName := NamespaceName,
		sourceClassName := ClassName,
		sourcePOUName := __POUNAME(),
		sourcePosition := __POSITION(),
		sourceDataType := TypeClass,
		targetDataType := GENERIC_TYPE_CLASS.UINT_16
	);
END_METHOD

(*!
<summary>Formats a supported generic value as text with capacity for 255 characters.</summary>
<description>
Requires live storage matching the descriptor. Same-encoding string values are copied directly into the
result, retaining at most 255 code units and a terminator without an intermediate 80-character string. STRING
input is converted directly into the result with STRING_TO_WSTRING2, using the library single-byte string
conversion rather than UTF-8 decoding. Output is truncated to 255 wide code units when needed; the function
completion flag is intentionally ignored because this API permits truncation. Numeric formatting retains its
native conversion behavior. Unsupported conversions raise GenericConversionNotSupportedException; the source
and ownership are unchanged. Descendants cannot override this descriptor operation; customize value equality
through IEqualityComparer or the stored object equality contract.
</description>
*)
METHOD FINAL AsWString255 : WSTRING(255)
VAR
	universalPointer : UNIVERSAL_POINTER;
END_VAR
universalPointer.AsByte := Address;

CASE TypeClass OF
	GENERIC_TYPE_CLASS.BOOLEAN:
		 AsWString255 := TO_WSTRING(universalPointer.AsBool^);
		 RETURN;
    GENERIC_TYPE_CLASS.INT_8:
		 AsWString255 := TO_WSTRING(universalPointer.AsSInt^);
		 RETURN;
    GENERIC_TYPE_CLASS.INT_16:
		 AsWString255 := TO_WSTRING(universalPointer.AsInt^);
		 RETURN;
    GENERIC_TYPE_CLASS.INT_32:
		 AsWString255 := TO_WSTRING(universalPointer.AsDInt^);
		 RETURN;
    GENERIC_TYPE_CLASS.INT_64:
		 AsWString255 := TO_WSTRING(universalPointer.AsLInt^);
		 RETURN;
    GENERIC_TYPE_CLASS.UINT_8:
		 AsWString255 := TO_WSTRING(universalPointer.AsUSInt^);
		 RETURN;
    GENERIC_TYPE_CLASS.UINT_16:
		 AsWString255 := TO_WSTRING(universalPointer.AsUInt^);
		 RETURN;
    GENERIC_TYPE_CLASS.UINT_32:
		 AsWString255 := TO_WSTRING(universalPointer.AsUDInt^);
		 RETURN;
    GENERIC_TYPE_CLASS.UINT_64:
		 AsWString255 := TO_WSTRING(universalPointer.AsULInt^);
		 RETURN;
    GENERIC_TYPE_CLASS.REAL_32:
		 AsWString255 := TO_WSTRING(universalPointer.AsReal^);
		 RETURN;
    GENERIC_TYPE_CLASS.REAL_64:
		 AsWString255 := TO_WSTRING(universalPointer.AsLReal^);
		 RETURN;
    GENERIC_TYPE_CLASS.STRING_8:
		Tc2_Utilities.STRING_TO_WSTRING2(
			pDstWSTRING := ADR(AsWString255),
			pSrcSTRING := universalPointer.AsString,
			nDstSize := SIZEOF(AsWString255)
		);
		 RETURN;
	GENERIC_TYPE_CLASS.STRING_16:
		Tc2_Utilities.WSTRNCPY(
			pDst := ADR(AsWString255),
			pSrc := universalPointer.AsWString,
			nDstSize := SIZEOF(AsWString255)
		);
		 RETURN;
    GENERIC_TYPE_CLASS.TIME_32:
		 AsWString255 := TO_WSTRING(universalPointer.AsTime^);
		 RETURN;
    GENERIC_TYPE_CLASS.TIME_64:
		 AsWString255 := TO_WSTRING(universalPointer.AsLTime^);
		 RETURN;
    GENERIC_TYPE_CLASS.DATE_32:
		 AsWString255 := TO_WSTRING(universalPointer.AsDate^);
		 RETURN;
    GENERIC_TYPE_CLASS.DATE_64:
		 AsWString255 := TO_WSTRING(universalPointer.AsLDate^);
		 RETURN;
    GENERIC_TYPE_CLASS.DATE_AND_TIME_32:
		 AsWString255 := TO_WSTRING(universalPointer.AsDateAndTime^);
		 RETURN;
    GENERIC_TYPE_CLASS.DATE_AND_TIME_64:
		 AsWString255 := TO_WSTRING(universalPointer.AsLDateAndTime^);
		 RETURN;
    GENERIC_TYPE_CLASS.TIME_OF_DAY_32:
		 AsWString255 := TO_WSTRING(universalPointer.AsTimeOfDay^);
		 RETURN;
    GENERIC_TYPE_CLASS.TIME_OF_DAY_64:
		 AsWString255 := TO_WSTRING(universalPointer.AsLTimeOfDay^);
		 RETURN;
END_CASE

Exceptions.ThrowGenericConversionNotSupported(
		sourceNamespaceName := NamespaceName,
		sourceClassName := ClassName,
		sourcePOUName := __POUNAME(),
		sourcePosition := __POSITION(),
		sourceDataType := TypeClass,
		targetDataType := GENERIC_TYPE_CLASS.STRING_16
	);
END_METHOD

(*!
<summary>Borrows the WSTRING storage described by this value.</summary>
<description>
Requires STRING_16 or raises GenericConversionNotSupportedException. Does not copy, bound-check or validate
the payload. The reference remains valid only while the source storage remains alive; the descriptor size
still limits any access. Descendants cannot override this descriptor operation; customize value equality
through IEqualityComparer or the stored object equality contract.
</description>
*)
METHOD FINAL AsWStringReference : REFERENCE TO WSTRING
VAR
	universalPointer : UNIVERSAL_POINTER;
END_VAR
universalPointer.AsByte := Address;

CASE TypeClass OF
	GENERIC_TYPE_CLASS.STRING_16:
		 AsWStringReference REF= universalPointer.AsWString^;
		 RETURN;
END_CASE

Exceptions.ThrowGenericConversionNotSupported(
		sourceNamespaceName := NamespaceName,
		sourceClassName := ClassName,
		sourcePOUName := __POUNAME(),
		sourcePosition := __POSITION(),
		sourceDataType := TypeClass,
		targetDataType := GENERIC_TYPE_CLASS.STRING_16
	);
END_METHOD

(*!
<summary>Changes the stored value using an ANY descriptor.</summary>
<description>
Delegates to ChangeValueByAnyType with the supplied isObject flag. Its compatibility checks, ownership
behavior, mutation rules and exceptions apply unchanged; input storage is borrowed during the call.
Descendants cannot override this descriptor operation; customize value equality through IEqualityComparer or
the stored object equality contract.
</description>
*)
METHOD FINAL ChangeValueByAny
VAR_INPUT
	value : ANY;
	isObject : BOOL := FALSE;
END_VAR
ChangeValueByAnyType(value := value, isObject := isObject);
END_METHOD

(*!
<summary>Copies a compatible source into existing storage and reports validation or native copy failure.</summary>
<description>
Both descriptors must refer to live storage. Type and capacity are checked before writing. No allocation,
ownership transfer or descriptor mutation occurs. The caller handles native exceptions and partial writes.
</description>
<param name="value">Borrowed source descriptor.</param>
<param name="sourceType">Generic category already resolved for the source.</param>
*)
METHOD PRIVATE copyMappedValue : GENERIC_VALUE_COPY_RESULT
VAR_INPUT
	value : __SYSTEM.AnyType;
	sourceType : GENERIC_TYPE_CLASS;
END_VAR
IF sourceType <> TypeClass THEN
	copyMappedValue := GENERIC_VALUE_COPY_RESULT.INCOMPATIBLE_TYPE;
	RETURN;
END_IF

IF Size < TO_ULINT(value.diSize) THEN
	copyMappedValue := GENERIC_VALUE_COPY_RESULT.INSUFFICIENT_CAPACITY;
	RETURN;
END_IF

IF Tc2_System.MEMCPY(destAddr := Address, srcAddr := value.pValue, n := TO_UDINT(value.diSize)) = 0 THEN
	copyMappedValue := GENERIC_VALUE_COPY_RESULT.COPY_FAILED;
	RETURN;
END_IF

copyMappedValue := GENERIC_VALUE_COPY_RESULT.COPIED;
END_METHOD

(*!
<summary>Copies bytes from an AnyType value into the existing generic storage.</summary>
<description>
Maps the source type using isObject, then rejects a mismatched generic type through
IncompatibleGenericValueTypeException or insufficient destination capacity through
TargetVariableMemoryOverflowException. Copies value.diSize bytes with MEMCPY; a zero return raises
StandardException. Source type mapping exceptions propagate. Successful copying does not allocate, clone objects, change
descriptor fields or transfer ownership; bytes beyond the copied region remain unchanged. The caller supplies
valid descriptors and live storage; this method does not validate memory lifetime or guarantee
overlapping-copy behavior. Descendants cannot override this descriptor operation; customize value equality
through IEqualityComparer or the stored object equality contract.
</description>
*)
METHOD FINAL ChangeValueByAnyType
VAR_INPUT
	value : __SYSTEM.AnyType;
	isObject : BOOL := FALSE;
END_VAR
VAR
	argumentDataType : GENERIC_TYPE_CLASS;
END_VAR
argumentDataType := GenericTypeClassConvertor.GetGenericTypeClassBySystemAnyType(
	systemAnyType := value,
	isObject := isObject
);

CASE copyMappedValue(value := value, sourceType := argumentDataType) OF
	GENERIC_VALUE_COPY_RESULT.INCOMPATIBLE_TYPE:
		Exceptions.ThrowIncompatibleGenericValueType(
			sourceNamespaceName := NamespaceName,
			sourceClassName := ClassName,
			sourcePOUName := __POUNAME(),
			sourcePosition := __POSITION(),
			validatedObjectName := "value",
			actualTypeClass := argumentDataType,
			expectedTypeClass := TypeClass
		);

	GENERIC_VALUE_COPY_RESULT.INSUFFICIENT_CAPACITY:
		Exceptions.ThrowTargetVariableMemoryOverflow(
			sourceNamespaceName := NamespaceName,
			sourceClassName := ClassName,
			sourcePOUName := __POUNAME(),
			sourcePosition := __POSITION(),
			targetVariableName := 'Size',
			targetVariableSize := Size
		);

	GENERIC_VALUE_COPY_RESULT.COPY_FAILED:
		Exceptions.ThrowStandard(
			sourceNamespaceName := NamespaceName,
			sourceClassName := ClassName,
			sourcePOUName := __POUNAME(),
			sourcePosition := __POSITION(),
			message := "Tc2_System.MEMCPY returned error (value 0)"
		);
END_CASE
END_METHOD

{attribute 'monitoring' := 'call'}
PROPERTY ClassName : REFERENCE TO STRING
GET
ClassName REF= GenericValueFactory.GenericValueClassName;
END_GET
END_PROPERTY

(*!
<summary>Compares an integer descriptor with a non-NaN binary64 value without rounding the integer.</summary>
<description>
Requires live BOOLEAN or integer storage and the binary64 bits returned by getCanonicalRealBits for a non-NaN
REAL or LREAL. Does not allocate or convert the integer to floating-point. Separates signs, compares unsigned
magnitudes and reverses the result when both operands are negative. Handles signed minimum, negative zero,
fractions, subnormal values and infinities. The masks apply to binary64 storage; no NaN arithmetic is used.
</description>
<param name="integerValue">Borrowed BOOLEAN or integer descriptor.</param>
<param name="realBits">Non-NaN binary64 representation, with either signed zero representation allowed.</param>
*)
METHOD PRIVATE compareIntegerToReal : COMPARISON_RESULT
VAR_INPUT
	integerValue : GENERIC_VALUE;
	realBits : ULINT;
END_VAR
VAR CONSTANT
	//! <summary>Bias subtracted from the stored binary64 exponent to obtain its power of two.</summary>
	EXPONENT_BIAS : UINT := 1023;
	//! <summary>Number of stored binary64 fraction bits below the implicit leading bit.</summary>
	FRACTION_BIT_COUNT : UINT := 52;
	//! <summary>Width of the unsigned magnitude used to compare every supported integer representation.</summary>
	INTEGER_BIT_COUNT : UINT := SIZEOF(ULINT) * 8;
	//! <summary>Bit 52 restored above the stored binary64 fraction for a normal finite value.</summary>
	IMPLICIT_LEADING_BIT : ULINT := ULINT#16#0010000000000000;
END_VAR
VAR
	signedValue : LINT;
	integerMagnitude : ULINT;
	integerNegative : BOOL;
	realNegative : BOOL;
	realMagnitudeBits : ULINT;
	storedExponent : UINT;
	significand : ULINT;
	wholeMagnitude : ULINT;
	fractionBits : ULINT;
	rightShift : UINT;
END_VAR
IF integerValue.TypeClass >= GENERIC_TYPE_CLASS.INT_8
	AND_THEN integerValue.TypeClass <= GENERIC_TYPE_CLASS.INT_64
THEN
	signedValue := integerValue.AsLInt();
	integerNegative := signedValue < SignedInt64.ZERO;

	IF integerNegative THEN
		// Avoid negating LINT minimum directly.
		integerMagnitude := TO_ULINT(-(signedValue + 1)) + 1;
	ELSE
		integerMagnitude := TO_ULINT(signedValue);
	END_IF
ELSE
	integerMagnitude := integerValue.AsULInt();
END_IF

realMagnitudeBits := realBits AND LongReals.MAGNITUDE_MASK;
realNegative := realBits > LongReals.MAGNITUDE_MASK AND_THEN realMagnitudeBits <> LongReals.ZERO_BITS;

IF integerNegative <> realNegative THEN
	IF integerNegative THEN
		compareIntegerToReal := COMPARISON_RESULT.FIRST_LESS_THAN_SECOND;
	ELSE
		compareIntegerToReal := COMPARISON_RESULT.FIRST_GREATER_THAN_SECOND;
	END_IF

	RETURN;
END_IF

storedExponent := TO_UINT(SHR(realBits AND LongReals.EXPONENT_MASK, FRACTION_BIT_COUNT));

IF storedExponent < EXPONENT_BIAS THEN
	IF integerMagnitude > UnsignedInt64.MIN_VALUE THEN
		compareIntegerToReal := COMPARISON_RESULT.FIRST_GREATER_THAN_SECOND;
	ELSIF realMagnitudeBits = LongReals.ZERO_BITS THEN
		compareIntegerToReal := COMPARISON_RESULT.FIRST_EQUAL_TO_SECOND;
	ELSE
		compareIntegerToReal := COMPARISON_RESULT.FIRST_LESS_THAN_SECOND;
	END_IF
ELSIF storedExponent >= EXPONENT_BIAS + INTEGER_BIT_COUNT THEN
	// Every magnitude at least 2^64, including infinity, exceeds all supported integer magnitudes.
	compareIntegerToReal := COMPARISON_RESULT.FIRST_LESS_THAN_SECOND;
ELSE
	significand := (realBits AND LongReals.FRACTION_MASK) OR IMPLICIT_LEADING_BIT;

	IF storedExponent >= EXPONENT_BIAS + FRACTION_BIT_COUNT THEN
		wholeMagnitude := SHL(significand, storedExponent - EXPONENT_BIAS - FRACTION_BIT_COUNT);
	ELSE
		rightShift := EXPONENT_BIAS + FRACTION_BIT_COUNT - storedExponent;
		wholeMagnitude := SHR(significand, rightShift);
		// Isolate the discarded low significand bits to distinguish a fraction from an exact integer.
		fractionBits := significand AND (SHL(ULINT#1, rightShift) - 1);
	END_IF

	IF integerMagnitude < wholeMagnitude THEN
		compareIntegerToReal := COMPARISON_RESULT.FIRST_LESS_THAN_SECOND;
	ELSIF integerMagnitude > wholeMagnitude THEN
		compareIntegerToReal := COMPARISON_RESULT.FIRST_GREATER_THAN_SECOND;
	ELSIF fractionBits <> UnsignedInt64.MIN_VALUE THEN
		compareIntegerToReal := COMPARISON_RESULT.FIRST_LESS_THAN_SECOND;
	ELSE
		compareIntegerToReal := COMPARISON_RESULT.FIRST_EQUAL_TO_SECOND;
	END_IF
END_IF

IF integerNegative THEN
	CASE compareIntegerToReal OF
		COMPARISON_RESULT.FIRST_LESS_THAN_SECOND:
			compareIntegerToReal := COMPARISON_RESULT.FIRST_GREATER_THAN_SECOND;
		COMPARISON_RESULT.FIRST_GREATER_THAN_SECOND:
			compareIntegerToReal := COMPARISON_RESULT.FIRST_LESS_THAN_SECOND;
	END_CASE
END_IF
END_METHOD

(*!
<summary>Compares this generic value with another using an optional comparer or built-in ordering rules.</summary>
<description>
When comparer is supplied, Compare receives copies of both GENERIC_VALUE descriptors. The comparer and operands
are borrowed only for the call; no payload is copied or released. Without a comparer, built-in ordering applies:
null is less than non-null, and two null values are equal. Numeric values (integers, booleans, floating-point)
compare across signedness and widths: all NaN encodings compare equal and precede every non-NaN number.
NaN is classified before floating conversion. Other floating-point pairs compare as LREAL. Mixed integer and
floating-point pairs compare exactly by sign, integer magnitude and binary64 exponent/significand, without
rounding the integer to floating-point. Integer pairs compare by value across signed and unsigned
representations. Times compare as LTIME durations, dates
and datetimes compare as LDATE_AND_TIME. Strings compare their complete terminated sequences by code unit,
widening single-byte characters to WORD for mixed encodings without allocation or a 255-character limit.
OBJECT operands delegate to IComparable when implemented. Incompatible representations raise GenericConversionNotSupportedException.
</description>
*)
//!<param name="otherValue">Descriptor of the value to compare.</param>
//!<param name="comparer">Optional borrowed ordering strategy; zero selects built-in ordering.</param>
METHOD FINAL CompareTo : COMPARISON_RESULT
VAR_INPUT
	otherValue : GENERIC_VALUE;
	comparer : IComparer := 0;
END_VAR
VAR
	firstLReal : LREAL;
	secondLReal : LREAL;
	firstLInt : LINT;
	secondLInt : LINT;
	firstULInt : ULINT;
	secondULInt : ULINT;
	firstLTime : LTIME;
	secondLTime : LTIME;
	firstLDateTime : LDATE_AND_TIME;
	secondLDateTime : LDATE_AND_TIME;
	firstStringData : UNIVERSAL_POINTER;
	secondStringData : UNIVERSAL_POINTER;
	firstCharacter : WORD;
	secondCharacter : WORD;
	characterIndex : UDINT;
	firstObject : POINTER TO Object;
	secondObject : POINTER TO Object;
	firstComparable : IComparable;
	secondComparable : IComparable;
	isFirstNumeric : BOOL;
	isSecondNumeric : BOOL;
	isFirstFloat : BOOL;
	isSecondFloat : BOOL;
	isFirstNaN : BOOL;
	isSecondNaN : BOOL;
END_VAR
IF comparer <> 0 THEN
	CompareTo := comparer.Compare(first := THIS^, second := otherValue);
	RETURN;
END_IF

IF IsNull THEN
	IF otherValue.IsNull THEN
		CompareTo := COMPARISON_RESULT.FIRST_EQUAL_TO_SECOND;
	ELSE
		CompareTo := COMPARISON_RESULT.FIRST_LESS_THAN_SECOND;
	END_IF

	RETURN;
ELSIF otherValue.IsNull THEN
	CompareTo := COMPARISON_RESULT.FIRST_GREATER_THAN_SECOND;
	RETURN;
END_IF

isFirstNumeric := (TypeClass >= GENERIC_TYPE_CLASS.BOOLEAN AND_THEN TypeClass <= GENERIC_TYPE_CLASS.REAL_64);
isSecondNumeric := (otherValue.TypeClass >= GENERIC_TYPE_CLASS.BOOLEAN AND_THEN otherValue.TypeClass <= GENERIC_TYPE_CLASS.REAL_64);

IF isFirstNumeric AND_THEN isSecondNumeric THEN
	isFirstFloat := (TypeClass = GENERIC_TYPE_CLASS.REAL_32 OR_ELSE TypeClass = GENERIC_TYPE_CLASS.REAL_64);
	isSecondFloat := (otherValue.TypeClass = GENERIC_TYPE_CLASS.REAL_32 OR_ELSE otherValue.TypeClass = GENERIC_TYPE_CLASS.REAL_64);

	IF isFirstFloat OR_ELSE isSecondFloat THEN
		isFirstNaN := isFirstFloat AND_THEN getCanonicalRealBits() = LongReals.CANONICAL_NAN_BITS;
		isSecondNaN := isSecondFloat AND_THEN otherValue.getCanonicalRealBits() = LongReals.CANONICAL_NAN_BITS;

		IF isFirstNaN THEN
			IF isSecondNaN THEN
				CompareTo := COMPARISON_RESULT.FIRST_EQUAL_TO_SECOND;
			ELSE
				CompareTo := COMPARISON_RESULT.FIRST_LESS_THAN_SECOND;
			END_IF

			RETURN;
		ELSIF isSecondNaN THEN
			CompareTo := COMPARISON_RESULT.FIRST_GREATER_THAN_SECOND;
			RETURN;
		END_IF

		IF NOT isFirstFloat THEN
			CompareTo := compareIntegerToReal(integerValue := THIS^, realBits := otherValue.getCanonicalRealBits());
			RETURN;
		ELSIF NOT isSecondFloat THEN
			CASE compareIntegerToReal(integerValue := otherValue, realBits := getCanonicalRealBits()) OF
				COMPARISON_RESULT.FIRST_LESS_THAN_SECOND:
					CompareTo := COMPARISON_RESULT.FIRST_GREATER_THAN_SECOND;
				COMPARISON_RESULT.FIRST_EQUAL_TO_SECOND:
					CompareTo := COMPARISON_RESULT.FIRST_EQUAL_TO_SECOND;
				COMPARISON_RESULT.FIRST_GREATER_THAN_SECOND:
					CompareTo := COMPARISON_RESULT.FIRST_LESS_THAN_SECOND;
			END_CASE

			RETURN;
		END_IF

		firstLReal := AsLReal();
		secondLReal := otherValue.AsLReal();

		IF firstLReal < secondLReal THEN
			CompareTo := COMPARISON_RESULT.FIRST_LESS_THAN_SECOND;
		ELSIF firstLReal > secondLReal THEN
			CompareTo := COMPARISON_RESULT.FIRST_GREATER_THAN_SECOND;
		ELSE
			CompareTo := COMPARISON_RESULT.FIRST_EQUAL_TO_SECOND;
		END_IF

		RETURN;
	END_IF

	IF (TypeClass >= GENERIC_TYPE_CLASS.INT_8 AND_THEN TypeClass <= GENERIC_TYPE_CLASS.INT_64) THEN
		IF (otherValue.TypeClass >= GENERIC_TYPE_CLASS.INT_8 AND_THEN otherValue.TypeClass <= GENERIC_TYPE_CLASS.INT_64) THEN
			firstLInt := AsLInt();
			secondLInt := otherValue.AsLInt();

			IF firstLInt < secondLInt THEN
				CompareTo := COMPARISON_RESULT.FIRST_LESS_THAN_SECOND;
			ELSIF firstLInt > secondLInt THEN
				CompareTo := COMPARISON_RESULT.FIRST_GREATER_THAN_SECOND;
			ELSE
				CompareTo := COMPARISON_RESULT.FIRST_EQUAL_TO_SECOND;
			END_IF

			RETURN;
		ELSE
			firstLInt := AsLInt();

			IF firstLInt < SignedInt64.ZERO THEN
				CompareTo := COMPARISON_RESULT.FIRST_LESS_THAN_SECOND;
			ELSE
				secondULInt := otherValue.AsULInt();

				IF TO_ULINT(firstLInt) < secondULInt THEN
					CompareTo := COMPARISON_RESULT.FIRST_LESS_THAN_SECOND;
				ELSIF TO_ULINT(firstLInt) > secondULInt THEN
					CompareTo := COMPARISON_RESULT.FIRST_GREATER_THAN_SECOND;
				ELSE
					CompareTo := COMPARISON_RESULT.FIRST_EQUAL_TO_SECOND;
				END_IF
			END_IF

			RETURN;
		END_IF
	ELSE
		IF (otherValue.TypeClass >= GENERIC_TYPE_CLASS.INT_8 AND_THEN otherValue.TypeClass <= GENERIC_TYPE_CLASS.INT_64) THEN
			secondLInt := otherValue.AsLInt();

			IF secondLInt < SignedInt64.ZERO THEN
				CompareTo := COMPARISON_RESULT.FIRST_GREATER_THAN_SECOND;
			ELSE
				firstULInt := AsULInt();

				IF firstULInt < TO_ULINT(secondLInt) THEN
					CompareTo := COMPARISON_RESULT.FIRST_LESS_THAN_SECOND;
				ELSIF firstULInt > TO_ULINT(secondLInt) THEN
					CompareTo := COMPARISON_RESULT.FIRST_GREATER_THAN_SECOND;
				ELSE
					CompareTo := COMPARISON_RESULT.FIRST_EQUAL_TO_SECOND;
				END_IF
			END_IF

			RETURN;
		ELSE
			firstULInt := AsULInt();
			secondULInt := otherValue.AsULInt();

			IF firstULInt < secondULInt THEN
				CompareTo := COMPARISON_RESULT.FIRST_LESS_THAN_SECOND;
			ELSIF firstULInt > secondULInt THEN
				CompareTo := COMPARISON_RESULT.FIRST_GREATER_THAN_SECOND;
			ELSE
				CompareTo := COMPARISON_RESULT.FIRST_EQUAL_TO_SECOND;
			END_IF

			RETURN;
		END_IF
	END_IF
END_IF

IF (TypeClass = GENERIC_TYPE_CLASS.TIME_32 OR_ELSE TypeClass = GENERIC_TYPE_CLASS.TIME_64) AND_THEN
   (otherValue.TypeClass = GENERIC_TYPE_CLASS.TIME_32 OR_ELSE otherValue.TypeClass = GENERIC_TYPE_CLASS.TIME_64) THEN
	firstLTime := AsLTime();
	secondLTime := otherValue.AsLTime();

	IF firstLTime < secondLTime THEN
		CompareTo := COMPARISON_RESULT.FIRST_LESS_THAN_SECOND;
	ELSIF firstLTime > secondLTime THEN
		CompareTo := COMPARISON_RESULT.FIRST_GREATER_THAN_SECOND;
	ELSE
		CompareTo := COMPARISON_RESULT.FIRST_EQUAL_TO_SECOND;
	END_IF

	RETURN;
END_IF

IF (TypeClass = GENERIC_TYPE_CLASS.DATE_32 OR_ELSE TypeClass = GENERIC_TYPE_CLASS.DATE_64 OR_ELSE
    TypeClass = GENERIC_TYPE_CLASS.DATE_AND_TIME_32 OR_ELSE TypeClass = GENERIC_TYPE_CLASS.DATE_AND_TIME_64) AND_THEN
   (otherValue.TypeClass = GENERIC_TYPE_CLASS.DATE_32 OR_ELSE otherValue.TypeClass = GENERIC_TYPE_CLASS.DATE_64 OR_ELSE
    otherValue.TypeClass = GENERIC_TYPE_CLASS.DATE_AND_TIME_32 OR_ELSE otherValue.TypeClass = GENERIC_TYPE_CLASS.DATE_AND_TIME_64) THEN
	firstLDateTime := AsLDateAndTime();
	secondLDateTime := otherValue.AsLDateAndTime();

	IF firstLDateTime < secondLDateTime THEN
		CompareTo := COMPARISON_RESULT.FIRST_LESS_THAN_SECOND;
	ELSIF firstLDateTime > secondLDateTime THEN
		CompareTo := COMPARISON_RESULT.FIRST_GREATER_THAN_SECOND;
	ELSE
		CompareTo := COMPARISON_RESULT.FIRST_EQUAL_TO_SECOND;
	END_IF

	RETURN;
END_IF

IF (TypeClass = GENERIC_TYPE_CLASS.STRING_8 OR_ELSE TypeClass = GENERIC_TYPE_CLASS.STRING_16)
	AND_THEN (otherValue.TypeClass = GENERIC_TYPE_CLASS.STRING_8
		OR_ELSE otherValue.TypeClass = GENERIC_TYPE_CLASS.STRING_16)
THEN
	firstStringData.AsByte := Address;
	secondStringData.AsByte := otherValue.Address;

	WHILE TRUE DO
		IF TypeClass = GENERIC_TYPE_CLASS.STRING_8 THEN
			firstCharacter := TO_WORD(firstStringData.AsByte[characterIndex]);
		ELSE
			firstCharacter := firstStringData.AsWord[characterIndex];
		END_IF

		IF otherValue.TypeClass = GENERIC_TYPE_CLASS.STRING_8 THEN
			secondCharacter := TO_WORD(secondStringData.AsByte[characterIndex]);
		ELSE
			secondCharacter := secondStringData.AsWord[characterIndex];
		END_IF

		IF firstCharacter < secondCharacter THEN
			CompareTo := COMPARISON_RESULT.FIRST_LESS_THAN_SECOND;
			RETURN;
		ELSIF firstCharacter > secondCharacter THEN
			CompareTo := COMPARISON_RESULT.FIRST_GREATER_THAN_SECOND;
			RETURN;
		ELSIF firstCharacter = TO_WORD(UnsignedInt16.MIN_VALUE) THEN
			CompareTo := COMPARISON_RESULT.FIRST_EQUAL_TO_SECOND;
			RETURN;
		END_IF

		characterIndex := characterIndex + 1;
	END_WHILE
END_IF

IF TypeClass = GENERIC_TYPE_CLASS.OBJECT AND_THEN otherValue.TypeClass = GENERIC_TYPE_CLASS.OBJECT THEN
	firstObject := Address;
	secondObject := otherValue.Address;
	
	IF __QUERYINTERFACE(firstObject^, firstComparable) AND_THEN __QUERYINTERFACE(secondObject^, secondComparable) THEN
		CompareTo := firstComparable.CompareTo(otherValue := secondComparable);
		RETURN;
	END_IF
END_IF

